   F[1631] := 3.685619;
   F[1632] := 3.6892362;
   F[1633] := 3.725405;
   F[1634] := 3.6639178;
   F[1635] := 3.6385996;
   F[1636] := 3.5879629;
   F[1637] := 3.6385996;
   F[1638] := 3.5807292;
   F[1639] := 3.59158;
   F[1640] := 3.5264757;
   F[1641] := 3.5083911;
   F[1642] := 3.5228589;
   F[1643] := 3.5300925;
   F[1644] := 3.4975405;
   F[1645] := 3.5011575;
   F[1646] := 3.4324362;
   F[1647] := 3.4252026;
   F[1648] := 3.5011575;
   F[1649] := 3.4324362;
   F[1650] := 3.410735;
   F[1651] := 3.4360533;
   F[1652] := 3.3962674;
   F[1653] := 3.374566;
   F[1654] := 3.370949;
   F[1655] := 3.3673322;
   F[1656] := 3.3528645;
   F[1657] := 3.3166957;
   F[1658] := 3.378183;
   F[1659] := 3.302228;
   F[1660] := 3.2841434;
   F[1661] := 3.294994;
   F[1662] := 3.233507;
   F[1663] := 3.2732928;
   F[1664] := 3.2045717;
   F[1665] := 3.226273;
   F[1666] := 3.1864872;
   F[1667] := 3.2045717;
   F[1668] := 3.2118056;
   F[1669] := 3.1394675;
   F[1670] := 3.157552;
   F[1671] := 3.161169;
   F[1672] := 3.1358507;
   F[1673] := 3.1286168;
   F[1674] := 3.1286168;
   F[1675] := 3.0454283;
   F[1676] := 3.0635128;
   F[1677] := 3.0996816;
   F[1678] := 3.0454283;
   F[1679] := 3.049045;
   F[1680] := 3.049045;
   F[1681] := 3.023727;
   F[1682] := 3.0092592;
   F[1683] := 2.9513888;
   F[1684] := 2.9513888;
   F[1685] := 2.983941;
   F[1686] := 2.980324;
   F[1687] := 2.9296875;
   F[1688] := 2.911603;
   F[1689] := 2.8573496;
   F[1690] := 2.8645833;
   F[1691] := 2.9188368;
   F[1692] := 2.911603;
   F[1693] := 2.8175638;
   F[1694] := 2.8537326;
   F[1695] := 2.842882;
   F[1696] := 2.8320312;
   F[1697] := 2.7958622;
   F[1698] := 2.7777777;
   F[1699] := 2.8139467;
   F[1700] := 2.734375;
   F[1701] := 2.7199075;
   F[1702] := 2.7596934;
   F[1703] := 2.7162905;
   F[1704] := 2.698206;
   F[1705] := 2.7416089;
   F[1706] := 2.6945891;
   F[1707] := 2.6801214;
   F[1708] := 2.6728878;
   F[1709] := 2.6367188;
   F[1710] := 2.629485;
   F[1711] := 2.6801214;
   F[1712] := 2.6367188;
   F[1713] := 2.6150174;
   F[1714] := 2.5752316;
   F[1715] := 2.564381;
   F[1716] := 2.55353;
   F[1717] := 2.5788484;
   F[1718] := 2.5426793;
   F[1719] := 2.4920428;
   F[1720] := 2.5282118;
   F[1721] := 2.5065105;
   F[1722] := 2.5028934;
   F[1723] := 2.4775753;
   F[1724] := 2.44864;
   F[1725] := 2.4088542;
   F[1726] := 2.4233217;
   F[1727] := 2.5065105;
   F[1728] := 2.3980036;
   F[1729] := 2.445023;
   F[1730] := 2.3582175;
   F[1731] := 2.4233217;
   F[1732] := 2.3618345;
   F[1733] := 2.376302;
   F[1734] := 2.3654513;
   F[1735] := 2.2858796;
   F[1736] := 2.3184316;
   F[1737] := 2.23886;
   F[1738] := 2.3365161;
   F[1739] := 2.275029;
   F[1740] := 2.2605612;
   F[1741] := 2.1918402;
   F[1742] := 2.2280092;
   F[1743] := 1.634838;
   F[1744] := 0.9765625;
   F[1745] := 0.30020255;
   F[1746] := 3.4432871;
   F[1747] := 5.0455728;
   F[1748] := 5.0998263;
   F[1749] := 5.10706;
   F[1750] := 5.0853586;
   F[1751] := 5.1613135;
   F[1752] := 5.117911;
   F[1753] := 5.128762;
   F[1754] := 5.0925927;
   F[1755] := 5.143229;
   F[1756] := 5.0600405;
   F[1757] := 5.0708914;
   F[1758] := 5.1649303;
   F[1759] := 5.128762;
   F[1760] := 5.114294;
   F[1761] := 5.103443;
   F[1762] := 5.1576967;
   F[1763] := 5.183015;
   F[1764] := 5.117911;
   F[1765] := 5.1576967;
   F[1766] := 5.179398;
   F[1767] := 5.1649303;
   F[1768] := 5.0708914;
   F[1769] := 5.1251445;
   F[1770] := 5.215567;
   F[1771] := 5.179398;
   F[1772] := 5.2119503;
   F[1773] := 5.1721644;
   F[1774] := 5.204716;
   F[1775] := 5.150463;
   F[1776] := 5.204716;
   F[1777] := 5.179398;
   F[1778] := 5.190249;
   F[1779] := 5.1974826;
   F[1780] := 5.2445025;
   F[1781] := 5.2408853;
   F[1782] := 5.1757812;
   F[1783] := 5.251736;
   F[1784] := 5.280671;
   F[1785] := 5.2445025;
   F[1786] := 5.255353;
   F[1787] := 5.2842884;
   F[1788] := 5.2408853;
   F[1789] := 5.280671;
   F[1790] := 5.2445025;
   F[1791] := 5.2336516;
   F[1792] := 5.2987556;
   F[1793] := 5.230035;
   F[1794] := 5.2698207;
   F[1795] := 5.31684;
   F[1796] := 5.3783274;
   F[1797] := 5.3385415;
   F[1798] := 5.2987556;
   F[1799] := 5.287905;
   F[1800] := 5.3132234;
   F[1801] := 5.2770543;
   F[1802] := 5.3747106;
   F[1803] := 5.3132234;
   F[1804] := 5.4000287;
   F[1805] := 5.353009;
   F[1806] := 5.3096066;
   F[1807] := 5.6315103;
   F[1808] := 6.3368053;
   F[1809] := 6.969763;
   F[1810] := 7.60272;
   F[1811] := 8.282697;
   F[1812] := 8.427373;
   F[1813] := 8.405671;
   F[1814] := 8.445457;
   F[1815] := 8.456307;
   F[1816] := 8.423756;
   F[1817] := 8.510561;
   F[1818] := 8.539496;
   F[1819] := 8.564815;
   F[1820] := 8.496094;
   F[1821] := 8.59375;
   F[1822] := 8.600984;
   F[1823] := 8.619068;
   F[1824] := 8.557581;
   F[1825] := 8.691406;
   F[1826] := 8.669704;
   F[1827] := 8.691406;
   F[1828] := 8.738426;
   F[1829] := 8.637153;
   F[1830] := 8.763744;
   F[1831] := 8.781829;
   F[1832] := 8.796296;
   F[1833] := 8.785445;
   F[1834] := 8.80353;
   F[1835] := 8.843316;
   F[1836] := 8.854167;
   F[1837] := 8.875868;
   F[1838] := 8.843316;
   F[1839] := 8.908421;
   F[1840] := 8.937355;
   F[1841] := 8.9192705;
   F[1842] := 9.006077;
   F[1843] := 8.959057;
   F[1844] := 8.998842;
   F[1845] := 8.973524;
   F[1846] := 9.016927;
   F[1847] := 9.031395;
   F[1848] := 9.031395;
   F[1849] := 8.998842;
   F[1850] := 9.085649;
   F[1851] := 9.063947;
   F[1852] := 9.154369;
   F[1853] := 9.186921;
   F[1854] := 9.161603;
   F[1855] := 9.273726;
   F[1856] := 9.201389;
   F[1857] := 9.226707;
   F[1858] := 9.233941;
   F[1859] := 9.248408;
   F[1860] := 9.248408;
   F[1861] := 9.338831;
   F[1862] := 9.338831;
   F[1863] := 9.349682;
   F[1864] := 9.302662;
   F[1865] := 9.364149;
   F[1866] := 9.447338;
   F[1867] := 9.367766;
   F[1868] := 9.454572;
   F[1869] := 9.385851;
   F[1870] := 9.42202;
   F[1871] := 9.476274;
   F[1872] := 9.490741;
   F[1873] := 9.505208;
   F[1874] := 9.505208;
   F[1875] := 9.602864;
   F[1876] := 9.555845;
   F[1877] := 9.544994;
   F[1878] := 9.588397;
   F[1879] := 9.628182;
   F[1880] := 9.664351;
   F[1881] := 9.628182;
   F[1882] := 9.660735;
   F[1883] := 9.682436;
   F[1884] := 9.729456;
   F[1885] := 9.707755;
   F[1886] := 9.73669;
   F[1887] := 9.740307;
   F[1888] := 9.823495;
   F[1889] := 9.805411;
   F[1890] := 9.798177;
   F[1891] := 9.823495;
   F[1892] := 9.866899;
   F[1893] := 9.881366;
   F[1894] := 9.85243;
   F[1895] := 9.975405;
   F[1896] := 10.007957;
   F[1897] := 9.95732;
   F[1898] := 10.029658;
   F[1899] := 10.185185;
   F[1900] := 10.206886;
   F[1901] := 10.315393;
   F[1902] := 10.467303;
   F[1903] := 10.554109;
   F[1904] := 10.691551;
   F[1905] := 10.756655;
   F[1906] := 10.789207;
   F[1907] := 10.966435;
   F[1908] := 11.067708;
   F[1909] := 11.161748;
   F[1910] := 11.205151;
   F[1911] := 11.338976;
   F[1912] := 11.472801;
   F[1913] := 11.555989;
   F[1914] := 11.603009;
   F[1915] := 11.715133;
   F[1916] := 11.794704;
   F[1917] := 11.924913;
   F[1918] := 12.040654;
   F[1919] := 12.131077;
   F[1920] := 12.203414;
   F[1921] := 12.355324;
   F[1922] := 12.384259;
   F[1923] := 12.507234;
   F[1924] := 12.60489;
   F[1925] := 12.648293;
   F[1926] := 12.800202;
   F[1927] := 12.9557295;
   F[1928] := 13.042535;
   F[1929] := 13.078704;
   F[1930] := 13.165509;
   F[1931] := 13.32827;
   F[1932] := 13.404224;
   F[1933] := 13.527199;
   F[1934] := 13.58507;
   F[1935] := 13.726129;
   F[1936] := 13.820168;
   F[1937] := 13.968461;
   F[1938] := 13.990162;
   F[1939] := 14.134838;
   F[1940] := 14.21441;
   F[1941] := 14.279514;
   F[1942] := 14.362702;
   F[1943] := 14.532697;
   F[1944] := 14.619502;
   F[1945] := 14.7316265;
   F[1946] := 14.840133;
   F[1947] := 14.923322;
   F[1948] := 14.623119;
   F[1949] := 13.798467;
   F[1950] := 12.9557295;
   F[1951] := 12.160011;
   F[1952] := 11.382379;
   F[1953] := 11.020689;
   F[1954] := 11.053241;
   F[1955] := 11.121962;
   F[1956] := 11.107494;
   F[1957] := 11.143663;
   F[1958] := 11.121962;
   F[1959] := 11.150897;
   F[1960] := 11.14728;
   F[1961] := 11.219618;
   F[1962] := 11.190682;
   F[1963] := 11.183449;
   F[1964] := 11.223235;
   F[1965] := 11.302807;
   F[1966] := 11.295573;
   F[1967] := 11.255787;
   F[1968] := 11.364294;
   F[1969] := 11.317274;
   F[1970] := 11.375145;
   F[1971] := 11.3932295;
   F[1972] := 11.418548;
   F[1973] := 11.4402485;
   F[1974] := 11.469184;
   F[1975] := 11.436632;
   F[1976] := 11.494502;
   F[1977] := 11.494502;
   F[1978] := 11.588542;
   F[1979] := 11.555989;
   F[1980] := 11.559607;
   F[1981] := 11.603009;
   F[1982] := 11.617476;
   F[1983] := 11.617476;
   F[1984] := 11.704283;
   F[1985] := 11.693432;
   F[1986] := 11.678964;
   F[1987] := 11.715133;
   F[1988] := 11.744068;
   F[1989] := 11.773004;
   F[1990] := 11.758536;
   F[1991] := 11.816406;
   F[1992] := 11.809173;
   F[1993] := 11.848958;
   F[1994] := 11.910445;
   F[1995] := 11.950232;
   F[1996] := 11.874276;
   F[1997] := 11.932147;
   F[1998] := 11.924913;
   F[1999] := 11.968316;
   F[2000] := 11.979167;
   F[2001] := 12.004485;
   F[2002] := 12.037037;
   F[2003] := 12.000868;
   F[2004] := 12.123842;
   F[2005] := 12.105758;
   F[2006] := 12.181713;
   F[2007] := 12.141927;
   F[2008] := 12.203414;
   F[2009] := 12.13831;
   F[2010] := 12.203414;
   F[2011] := 12.239583;
   F[2012] := 12.250434;
   F[2013] := 12.2432;
   F[2014] := 12.29022;
   F[2015] := 12.326389;
   F[2016] := 12.366175;
   F[2017] := 12.362557;
   F[2018] := 12.358941;
   F[2019] := 12.3878765;
   F[2020] := 12.3878765;
   F[2021] := 12.424046;
   F[2022] := 12.405961;
   F[2023] := 12.485533;
   F[2024] := 12.528935;
   F[2025] := 12.528935;
   F[2026] := 12.528935;
   F[2027] := 12.54702;
   F[2028] := 12.554254;
   F[2029] := 12.615741;
   F[2030] := 12.619358;
   F[2031] := 12.626592;
   F[2032] := 12.662761;
   F[2033] := 12.6953125;
   F[2034] := 12.764033;
   F[2035] := 12.811053;
   F[2036] := 12.724248;
   F[2037] := 12.760417;
   F[2038] := 12.80382;
   F[2039] := 12.843605;
   F[2040] := 12.836371;
   F[2041] := 12.850839;
   F[2042] := 12.90871;
   F[2043] := 12.941261;
   F[2044] := 13.292101;
   F[2045] := 15.704572;
   F[2046] := 18.17853;
   F[2047] := 20.706741;
   F[2048] := 23.1807;
   F[2049] := 25.672743;
   F[2050] := 28.121384;
   F[2051] := 30.671297;
   F[2052] := 33.15249;
   F[2053] := 35.633682;
   F[2054] := 38.151043;
   F[2055] := 40.588833;
   F[2056] := 40.559895;
   F[2057] := 37.492767;
   F[2058] := 34.964554;
   F[2059] := 32.508682;
   F[2060] := 30.016638;
   F[2061] := 27.50651;
   F[2062] := 25.043404;
   F[2063] := 22.518808;
   F[2064] := 20.070168;
   F[2065] := 17.520254;
   F[2066] := 15.089699;
   F[2067] := 12.579572;
   F[2068] := 11.237702;
   F[2069] := 11.161748;
   F[2070] := 11.2160015;
   F[2071] := 11.114728;
   F[2072] := 11.100261;
   F[2073] := 11.121962;
   F[2074] := 11.096643;
   F[2075] := 11.085793;
   F[2076] := 11.031539;
   F[2077] := 11.024305;
   F[2078] := 11.056858;
   F[2079] := 10.951967;
   F[2080] := 11.020689;
   F[2081] := 10.944734;
   F[2082] := 10.912182;
   F[2083] := 10.901331;
   F[2084] := 10.87963;
   F[2085] := 10.8253765;
   F[2086] := 10.803675;
   F[2087] := 10.789207;
   F[2088] := 10.73857;
   F[2089] := 10.745805;
   F[2090] := 10.781974;
   F[2091] := 10.706018;
   F[2092] := 10.724103;
   F[2093] := 10.593895;
   F[2094] := 10.673467;
   F[2095] := 10.6807;
   F[2096] := 10.572193;
   F[2097] := 10.554109;
   F[2098] := 10.579427;
   F[2099] := 10.503472;
   F[2100] := 10.521557;
   F[2101] := 10.52879;
   F[2102] := 10.463686;
   F[2103] := 10.445601;
   F[2104] := 10.46007;
   F[2105] := 10.532408;
   F[2106] := 10.420283;
   F[2107] := 10.35518;
   F[2108] := 10.322627;
   F[2109] := 10.326244;
   F[2110] := 10.3515625;
   F[2111] := 10.286458;
   F[2112] := 10.250289;
   F[2113] := 10.243055;
   F[2114] := 10.228588;
   F[2115] := 10.2213545;
   F[2116] := 10.181568;
   F[2117] := 10.206886;
   F[2118] := 10.192419;
   F[2119] := 10.083912;
   F[2120] := 10.112847;
   F[2121] := 10.083912;
   F[2122] := 10.054976;
   F[2123] := 10.047743;
   F[2124] := 10.007957;
   F[2125] := 10.007957;
   F[2126] := 9.964555;
   F[2127] := 9.982639;
   F[2128] := 9.986256;
   F[2129] := 9.924768;
   F[2130] := 9.89945;
   F[2131] := 9.892217;
   F[2132] := 9.848814;
   F[2133] := 9.837963;
   F[2134] := 9.884983;
   F[2135] := 9.801794;
   F[2136] := 9.780092;
   F[2137] := 9.780092;
   F[2138] := 9.754774;
   F[2139] := 9.725839;
   F[2140] := 9.725839;
   F[2141] := 9.711371;
   F[2142] := 9.693287;
   F[2143] := 9.6535015;
   F[2144] := 9.617332;
   F[2145] := 9.628182;
   F[2146] := 9.599248;
   F[2147] := 9.566695;
   F[2148] := 9.610099;
   F[2149] := 9.57393;
   F[2150] := 9.508825;
   F[2151] := 9.4871235;
   F[2152] := 9.443721;
   F[2153] := 9.414786;
   F[2154] := 9.43287;
   F[2155] := 9.382234;
   F[2156] := 9.382234;
   F[2157] := 9.360533;
   F[2158] := 9.324364;
   F[2159] := 9.338831;
   F[2160] := 9.306279;
   F[2161] := 9.378617;
   F[2162] := 9.244792;
   F[2163] := 9.215857;
   F[2164] := 9.2628765;
   F[2165] := 9.291811;
   F[2166] := 9.186921;
   F[2167] := 9.183305;
   F[2168] := 9.190538;
   F[2169] := 9.194155;
   F[2170] := 9.147136;
   F[2171] := 9.067564;
   F[2172] := 9.035011;
   F[2173] := 9.009693;
   F[2174] := 9.103733;
   F[2175] := 8.991609;
   F[2176] := 9.009693;
   F[2177] := 9.009693;
   F[2178] := 8.991609;
   F[2179] := 9.027778;
   F[2180] := 8.933739;
   F[2181] := 8.8722515;
   F[2182] := 8.933739;
   F[2183] := 8.865017;
   F[2184] := 8.875868;
   F[2185] := 8.843316;
   F[2186] := 8.7890625;
   F[2187] := 8.843316;
   F[2188] := 8.74566;
   F[2189] := 8.713108;
   F[2190] := 8.767361;
   F[2191] := 8.7058735;
   F[2192] := 8.687789;
   F[2193] := 8.673322;
   F[2194] := 8.7058735;
   F[2195] := 8.600984;
   F[2196] := 8.597367;
   F[2197] := 8.604601;
   F[2198] := 8.600984;
   F[2199] := 8.575665;
   F[2200] := 8.532263;
   F[2201] := 8.532263;
   F[2202] := 8.521412;
   F[2203] := 8.553964;
   F[2204] := 8.5286455;
   F[2205] := 8.478009;
   F[2206] := 8.4816265;
   F[2207] := 8.470776;
   F[2208] := 8.409288;
   F[2209] := 8.351418;
   F[2210] := 8.308015;
   F[2211] := 8.362268;
   F[2212] := 8.3152485;
   F[2213] := 8.3152485;
   F[2214] := 8.297164;
   F[2215] := 8.293548;
   F[2216] := 8.213976;
   F[2217] := 8.206742;
   F[2218] := 8.199508;
   F[2219] := 8.224827;
   F[2220] := 8.192274;
   F[2221] := 8.17419;
   F[2222] := 8.18504;
   F[2223] := 8.134404;
   F[2224] := 8.101851;
   F[2225] := 8.065682;
   F[2226] := 8.080151;
   F[2227] := 8.065682;
   F[2228] := 8.065682;
   F[2229] := 8.025897;
   F[2230] := 7.9716434;
   F[2231] := 8.036748;
   F[2232] := 7.9318576;
   F[2233] := 7.939091;
   F[2234] := 7.949942;
   F[2235] := 7.913773;
   F[2236] := 7.9029226;
   F[2237] := 7.8703704;
   F[2238] := 7.884838;
   F[2239] := 7.8956885;
   F[2240] := 7.837818;
   F[2241] := 7.8052664;
   F[2242] := 7.747396;
   F[2243] := 7.7582464;
   F[2244] := 7.7256947;
   F[2245] := 7.7546296;
   F[2246] := 7.703993;
   F[2247] := 7.6931424;
   F[2248] := 7.7293115;
   F[2249] := 7.6678243;
   F[2250] := 7.6171875;
   F[2251] := 7.5882525;
   F[2252] := 7.6497397;
   F[2253] := 7.5810184;
   F[2254] := 7.573785;
   F[2255] := 7.5810184;
   F[2256] := 7.530382;
   F[2257] := 7.5520835;
   F[2258] := 7.5050635;
   F[2259] := 7.486979;
   F[2260] := 7.472512;
   F[2261] := 7.5014467;
   F[2262] := 7.396557;
   F[2263] := 7.382089;
   F[2264] := 7.458044;
   F[2265] := 7.360388;
   F[2266] := 7.3423033;
   F[2267] := 7.349537;
   F[2268] := 7.309751;
   F[2269] := 7.3025174;
   F[2270] := 7.248264;
   F[2271] := 7.306134;
   F[2272] := 7.269965;
   F[2273] := 7.2265625;
   F[2274] := 7.1903934;
   F[2275] := 7.157841;
   F[2276] := 7.2012444;
   F[2277] := 7.139757;
   F[2278] := 7.168692;
   F[2279] := 7.1108217;
   F[2280] := 7.081887;
   F[2281] := 7.0746527;
   F[2282] := 7.0999713;
   F[2283] := 7.0457177;
   F[2284] := 7.1759257;
   F[2285] := 7.027633;
   F[2286] := 7.03125;
   F[2287] := 6.9878473;
   F[2288] := 6.9733796;
   F[2289] := 7.0131655;
   F[2290] := 6.929977;
   F[2291] := 6.8757234;
   F[2292] := 6.8974247;
   F[2293] := 6.857639;
   F[2294] := 6.8467884;
   F[2295] := 6.8865743;
   F[2296] := 6.8106194;
   F[2297] := 6.7599826;
   F[2298] := 6.792535;
   F[2299] := 6.814236;
   F[2300] := 6.792535;
   F[2301] := 6.2970195;
   F[2302] := 5.6351275;
   F[2303] := 4.875579;
   F[2304] := 4.257089;
   F[2305] := 3.6639178;
   F[2306] := 3.7073207;
   F[2307] := 3.69647;
   F[2308] := 3.6385996;
   F[2309] := 3.692853;
   F[2310] := 3.685619;
   F[2311] := 3.660301;
   F[2312] := 3.6639178;
   F[2313] := 3.6385996;
   F[2314] := 3.656684;
   F[2315] := 3.7181714;
   F[2316] := 3.685619;
   F[2317] := 3.6422164;
   F[2318] := 3.6277487;
   F[2319] := 3.620515;
   F[2320] := 3.6458333;
   F[2321] := 3.6385996;
   F[2322] := 3.5951967;
   F[2323] := 3.584346;
   F[2324] := 3.6313658;
   F[2325] := 3.5988138;
   F[2326] := 3.5879629;
   F[2327] := 3.5807292;
   F[2328] := 3.5879629;
   F[2329] := 3.5554109;
   F[2330] := 3.5879629;
   F[2331] := 3.59158;
   F[2332] := 3.551794;
   F[2333] := 3.5300925;
   F[2334] := 3.6060474;
   F[2335] := 3.5554109;
   F[2336] := 3.5300925;
   F[2337] := 3.5409434;
   F[2338] := 3.5264757;
   F[2339] := 3.5047743;
   F[2340] := 3.5192418;
   F[2341] := 3.5083911;
   F[2342] := 3.5373263;
   F[2343] := 3.5626447;
   F[2344] := 3.5011575;
   F[2345] := 3.5409434;
   F[2346] := 3.4866898;
   F[2347] := 3.5662615;
   F[2348] := 3.5120082;
   F[2349] := 3.5047743;
   F[2350] := 3.5192418;
   F[2351] := 3.4903066;
   F[2352] := 3.5228589;
   F[2353] := 3.4866898;
   F[2354] := 3.4505208;
   F[2355] := 3.4722223;
   F[2356] := 3.4649885;
   F[2357] := 3.446904;
   F[2358] := 3.4577546;
   F[2359] := 3.3528645;
   F[2360] := 3.4939237;
   F[2361] := 3.4866898;
   F[2362] := 3.4179688;
   F[2363] := 3.4215856;
   F[2364] := 3.4252026;
   F[2365] := 3.378183;
   F[2366] := 1.8916377;
   F[2367] := 4.615162;
   F[2368] := 4.626013;
   F[2369] := 4.5645256;
   F[2370] := 4.6187787;
   F[2371] := 4.6187787;
   F[2372] := 4.560909;
   F[2373] := 4.662182;
   F[2374] := 4.6296296;
   F[2375] := 4.6187787;
   F[2376] := 4.615162;
   F[2377] := 4.5645256;
   F[2378] := 4.622396;
   F[2379] := 4.6079283;
   F[2380] := 4.658565;
   F[2381] := 4.683883;
   F[2382] := 4.622396;
   F[2383] := 4.6043115;
   F[2384] := 4.691117;
   F[2385] := 4.6875;
   F[2386] := 4.676649;
   F[2387] := 4.647714;
   F[2388] := 4.6440973;
   F[2389] := 4.651331;
   F[2390] := 4.691117;
   F[2391] := 4.5898438;
   F[2392] := 4.6043115;
   F[2393] := 4.6730323;
   F[2394] := 4.723669;
   F[2395] := 4.6332464;
   F[2396] := 4.6730323;
   F[2397] := 4.7019677;
   F[2398] := 4.727286;
   F[2399] := 4.698351;
   F[2400] := 4.7019677;
   F[2401] := 4.6875;
   F[2402] := 4.6802664;
   F[2403] := 4.6730323;
   F[2404] := 4.6802664;
   F[2405] := 4.716435;
   F[2406] := 4.6947336;
   F[2407] := 4.6549478;
   F[2408] := 4.727286;
   F[2409] := 4.7345195;
   F[2410] := 4.738137;
   F[2411] := 4.727286;
   F[2412] := 4.788773;
   F[2413] := 4.7815394;
   F[2414] := 4.788773;
   F[2415] := 4.7670717;
   F[2416] := 4.7706885;
   F[2417] := 4.799624;
   F[2418] := 4.738137;
   F[2419] := 4.738137;
   F[2420] := 4.8177085;
   F[2421] := 4.763455;
   F[2422] := 4.8574944;
   F[2423] := 4.7815394;
   F[2424] := 4.7670717;
   F[2425] := 4.796007;
   F[2426] := 4.803241;
   F[2427] := 4.9479165;
   F[2428] := 5.5917244;
   F[2429] := 6.2934027;
   F[2430] := 6.919126;
   F[2431] := 7.526765;
   F[2432] := 7.8956885;
   F[2433] := 7.8920717;
   F[2434] := 7.8920717;
   F[2435] := 7.939091;
   F[2436] := 7.9029226;
   F[2437] := 7.960793;
   F[2438] := 7.960793;
   F[2439] := 7.960793;
   F[2440] := 7.9788775;
   F[2441] := 7.96441;
   F[2442] := 7.9463253;
   F[2443] := 8.036748;
   F[2444] := 8.018663;
   F[2445] := 8.087384;
   F[2446] := 8.065682;
   F[2447] := 8.105469;
   F[2448] := 8.141638;
   F[2449] := 8.188658;
   F[2450] := 8.145255;
   F[2451] := 8.181423;
   F[2452] := 8.192274;
   F[2453] := 8.17419;
   F[2454] := 8.275463;
   F[2455] := 8.206742;
   F[2456] := 8.199508;
   F[2457] := 8.308015;
   F[2458] := 8.257379;
   F[2459] := 8.311632;
   F[2460] := 8.326099;
   F[2461] := 8.33695;
   F[2462] := 8.322483;
   F[2463] := 8.33695;
   F[2464] := 8.3152485;
   F[2465] := 8.412905;
   F[2466] := 8.380353;
   F[2467] := 8.344184;
   F[2468] := 8.463542;
   F[2469] := 8.412905;
   F[2470] := 8.467158;
   F[2471] := 8.459925;
   F[2472] := 8.525029;
   F[2473] := 8.496094;
   F[2474] := 8.499711;
   F[2475] := 8.568432;
   F[2476] := 8.499711;
   F[2477] := 8.575665;
   F[2478] := 8.564815;
   F[2479] := 8.619068;
   F[2480] := 8.626302;
   F[2481] := 8.684173;
   F[2482] := 8.629919;
   F[2483] := 8.684173;
   F[2484] := 8.69864;
   F[2485] := 8.662471;
   F[2486] := 8.713108;
   F[2487] := 8.716724;
   F[2488] := 8.785445;
   F[2489] := 8.774595;
   F[2490] := 8.785445;
   F[2491] := 8.7890625;
   F[2492] := 8.79268;
   F[2493] := 8.846932;
   F[2494] := 8.825232;
   F[2495] := 8.904803;
   F[2496] := 8.890336;
   F[2497] := 8.930121;
   F[2498] := 8.987992;
   F[2499] := 8.973524;
   F[2500] := 8.944589;
   F[2501] := 8.933739;
   F[2502] := 9.07118;
   F[2503] := 9.01331;
   F[2504] := 9.038629;
   F[2505] := 9.020544;
   F[2506] := 9.056713;
   F[2507] := 9.07118;
   F[2508] := 9.038629;
   F[2509] := 9.125434;
   F[2510] := 9.1182;
   F[2511] := 9.103733;
   F[2512] := 9.190538;
   F[2513] := 9.139901;
   F[2514] := 9.215857;
   F[2515] := 9.244792;
   F[2516] := 9.226707;
   F[2517] := 9.284577;
   F[2518] := 9.302662;
   F[2519] := 9.400318;
   F[2520] := 9.519676;
   F[2521] := 9.602864;
   F[2522] := 9.696904;
   F[2523] := 9.801794;
   F[2524] := 9.870515;
   F[2525] := 9.94647;
   F[2526] := 10.058594;
   F[2527] := 10.174335;
   F[2528] := 10.275608;
   F[2529] := 10.380498;
   F[2530] := 10.456452;
   F[2531] := 10.568577;
   F[2532] := 10.698785;
   F[2533] := 10.745805;
   F[2534] := 10.836226;
   F[2535] := 10.944734;
   F[2536] := 11.078559;
   F[2537] := 11.085793;
   F[2538] := 11.248553;
   F[2539] := 11.367911;
   F[2540] := 11.458333;
   F[2541] := 11.530671;
   F[2542] := 11.621094;
   F[2543] := 11.700665;
   F[2544] := 11.841724;
   F[2545] := 11.92853;
   F[2546] := 12.029803;
   F[2547] := 12.152778;
   F[2548] := 12.207031;
   F[2549] := 12.344474;
   F[2550] := 12.377026;
   F[2551] := 12.518085;
   F[2552] := 12.637443;
   F[2553] := 12.713397;
   F[2554] := 12.811053;
   F[2555] := 12.883391;
   F[2556] := 13.064236;
   F[2557] := 13.089555;
   F[2558] := 13.22338;
   F[2559] := 13.292101;
   F[2560] := 13.436776;
   F[2561] := 13.527199;
   F[2562] := 13.610388;
   F[2563] := 13.718895;
   F[2564] := 13.820168;
   F[2565] := 13.932292;
   F[2566] := 14.001013;
   F[2567] := 14.073351;
   F[2568] := 13.943142;
   F[2569] := 13.136574;
   F[2570] := 12.380642;
   F[2571] := 11.563224;
   F[2572] := 10.662616;
   F[2573] := 10.199653;
   F[2574] := 10.206886;
   F[2575] := 10.275608;
   F[2576] := 10.264757;
   F[2577] := 10.257524;
   F[2578] := 10.271991;
   F[2579] := 10.282842;
   F[2580] := 10.322627;
   F[2581] := 10.402199;
   F[2582] := 10.3515625;
   F[2583] := 10.36603;
   F[2584] := 10.423901;
   F[2585] := 10.470921;
   F[2586] := 10.489005;
   F[2587] := 10.478154;
   F[2588] := 10.536024;
   F[2589] := 10.525173;
   F[2590] := 10.521557;
   F[2591] := 10.539641;
   F[2592] := 10.568577;
   F[2593] := 10.622829;
   F[2594] := 10.604745;
   F[2595] := 10.640914;
   F[2596] := 10.63368;
   F[2597] := 10.615596;
   F[2598] := 10.6589985;
   F[2599] := 10.698785;
   F[2600] := 10.767506;
   F[2601] := 10.687934;
   F[2602] := 10.724103;
   F[2603] := 10.78559;
   F[2604] := 10.807292;
   F[2605] := 10.854311;
   F[2606] := 10.756655;
   F[2607] := 10.821759;
   F[2608] := 10.774739;
   F[2609] := 10.876013;
   F[2610] := 10.857928;
   F[2611] := 10.894097;
   F[2612] := 10.857928;
   F[2613] := 10.926649;
   F[2614] := 10.930266;
   F[2615] := 10.988136;
   F[2616] := 11.035156;
   F[2617] := 11.046007;
   F[2618] := 11.038774;
   F[2619] := 11.017072;
   F[2620] := 11.096643;
   F[2621] := 11.118345;
   F[2622] := 11.085793;
   F[2623] := 11.143663;
   F[2624] := 11.201533;
   F[2625] := 11.1943;
   F[2626] := 11.201533;
   F[2627] := 11.176215;
   F[2628] := 11.230469;
   F[2629] := 11.205151;
   F[2630] := 11.342592;
   F[2631] := 11.291956;
   F[2632] := 11.31004;
   F[2633] := 11.313658;
   F[2634] := 11.313658;
   F[2635] := 11.331742;
   F[2636] := 11.41493;
   F[2637] := 11.443866;
   F[2638] := 11.407697;
   F[2639] := 11.46195;
   F[2640] := 11.447483;
   F[2641] := 11.490886;
   F[2642] := 11.51982;
   F[2643] := 11.541522;
   F[2644] := 11.545139;
   F[2645] := 11.501736;
   F[2646] := 11.628327;
   F[2647] := 11.621094;
   F[2648] := 11.628327;
   F[2649] := 11.639178;
   F[2650] := 11.624711;
   F[2651] := 11.646412;
   F[2652] := 11.682581;
   F[2653] := 11.729601;
   F[2654] := 11.71875;
   F[2655] := 11.791088;
   F[2656] := 11.794704;
   F[2657] := 11.856193;
   F[2658] := 11.834491;
   F[2659] := 11.780237;
   F[2660] := 11.845342;
   F[2661] := 11.852575;
   F[2662] := 11.859809;
   F[2663] := 11.932147;
   F[2664] := 12.084057;
   F[2665] := 14.369936;
   F[2666] := 16.880064;
   F[2667] := 19.382957;
   F[2668] := 21.849682;
   F[2669] := 24.374277;
   F[2670] := 26.837385;
   F[2671] := 29.394531;
   F[2672] := 31.807003;
   F[2673] := 34.324364;
   F[2674] := 36.816406;
   F[2675] := 39.304832;
   F[2676] := 41.82581;
   F[2677] := 41.822193;
   F[2678] := 38.697193;
   F[2679] := 36.23047;
   F[2680] := 33.716724;
   F[2681] := 31.210215;
   F[2682] := 28.68562;
   F[2683] := 26.182726;
   F[2684] := 23.672598;
   F[2685] := 21.216724;
   F[2686] := 18.75;
   F[2687] := 16.26519;
   F[2688] := 13.75868;
   F[2689] := 11.2160015;
   F[2690] := 10.21412;
   F[2691] := 10.170717;
   F[2692] := 10.199653;
   F[2693] := 10.116464;
   F[2694] := 10.058594;
   F[2695] := 10.112847;
   F[2696] := 10.073061;
   F[2697] := 10.10923;
   F[2698] := 10.080296;
   F[2699] := 9.993489;
   F[2700] := 10.015191;
   F[2701] := 10.040509;
   F[2702] := 9.968171;
   F[2703] := 9.928386;
   F[2704] := 9.924768;
   F[2705] := 9.982639;
   F[2706] := 9.942853;
   F[2707] := 9.859664;
   F[2708] := 9.870515;
   F[2709] := 9.845197;
   F[2710] := 9.845197;
   F[2711] := 9.834346;
   F[2712] := 9.85243;
   F[2713] := 9.686053;
   F[2714] := 9.765625;
   F[2715] := 9.725839;
   F[2716] := 9.73669;
   F[2717] := 9.718605;
   F[2718] := 9.7005205;
   F[2719] := 9.671586;
   F[2720] := 9.628182;
   F[2721] := 9.613715;
   F[2722] := 9.599248;
   F[2723] := 9.508825;
   F[2724] := 9.519676;
   F[2725] := 9.508825;
   F[2726] := 9.47989;
   F[2727] := 9.530526;
   F[2728] := 9.505208;
   F[2729] := 9.4401045;
   F[2730] := 9.461805;
   F[2731] := 9.458189;
   F[2732] := 9.396702;
   F[2733] := 9.360533;
   F[2734] := 9.389467;
   F[2735] := 9.295428;
   F[2736] := 9.331597;
   F[2737] := 9.306279;
   F[2738] := 9.284577;
   F[2739] := 9.313513;
   F[2740] := 9.233941;
   F[2741] := 9.295428;
   F[2742] := 9.230324;
   F[2743] := 9.226707;
   F[2744] := 9.215857;
   F[2745] := 9.136285;
   F[2746] := 9.129051;
   F[2747] := 9.0964985;
   F[2748] := 9.1182;
   F[2749] := 9.0964985;
   F[2750] := 9.056713;
   F[2751] := 9.085649;
   F[2752] := 9.042245;
   F[2753] := 9.016927;
   F[2754] := 8.998842;
   F[2755] := 9.006077;
   F[2756] := 8.959057;
   F[2757] := 8.995226;
   F[2758] := 8.933739;
   F[2759] := 8.886719;
   F[2760] := 8.868634;
   F[2761] := 8.868634;
   F[2762] := 8.886719;
   F[2763] := 8.861401;
   F[2764] := 8.825232;
   F[2765] := 8.846932;
   F[2766] := 8.723958;
   F[2767] := 8.7890625;
   F[2768] := 8.74566;
   F[2769] := 8.716724;
   F[2770] := 8.676939;
   F[2771] := 8.64077;
   F[2772] := 8.695024;
   F[2773] := 8.65162;
   F[2774] := 8.637153;
   F[2775] := 8.648004;
   F[2776] := 8.64077;
   F[2777] := 8.615452;
   F[2778] := 8.586516;
   F[2779] := 8.568432;
   F[2780] := 8.539496;
   F[2781] := 8.539496;
   F[2782] := 8.470776;
   F[2783] := 8.532263;
   F[2784] := 8.423756;
   F[2785] := 8.430989;
   F[2786] := 8.44184;
   F[2787] := 8.365886;
   F[2788] := 8.485243;
   F[2789] := 8.344184;
   F[2790] := 8.373119;
   F[2791] := 8.304399;
   F[2792] := 8.355035;
   F[2793] := 8.3152485;
   F[2794] := 8.300781;
   F[2795] := 8.246528;
   F[2796] := 8.297164;
   F[2797] := 8.257379;
   F[2798] := 8.235677;
   F[2799] := 8.206742;
   F[2800] := 8.199508;
   F[2801] := 8.177807;
   F[2802] := 8.159722;
   F[2803] := 8.152489;
   F[2804] := 8.065682;
   F[2805] := 8.148871;
   F[2806] := 8.083767;
   F[2807] := 8.065682;
   F[2808] := 8.051215;
   F[2809] := 8.047599;
   F[2810] := 8.029514;
   F[2811] := 8.01143;
   F[2812] := 7.9824944;
   F[2813] := 7.9571757;
   F[2814] := 7.9427085;
   F[2815] := 7.921007;
   F[2816] := 7.924624;
   F[2817] := 7.888455;
   F[2818] := 7.8956885;
   F[2819] := 7.8450522;
   F[2820] := 7.816117;
   F[2821] := 7.8305845;
   F[2822] := 7.873987;
   F[2823] := 7.7944155;
   F[2824] := 7.7980323;
   F[2825] := 7.675058;
   F[2826] := 7.751013;
   F[2827] := 7.736545;
   F[2828] := 7.675058;
   F[2829] := 7.6569734;
   F[2830] := 7.7329283;
   F[2831] := 7.664207;
   F[2832] := 7.6822915;
   F[2833] := 7.624421;
   F[2834] := 7.624421;
   F[2835] := 7.599103;
   F[2836] := 7.5810184;
   F[2837] := 7.5774016;
   F[2838] := 7.533999;
   F[2839] := 7.494213;
   F[2840] := 7.548466;
   F[2841] := 7.4652777;
   F[2842] := 7.530382;
   F[2843] := 7.4905963;
   F[2844] := 7.3893228;
   F[2845] := 7.411024;
   F[2846] := 7.3676214;
   F[2847] := 7.458044;
   F[2848] := 7.411024;
   F[2849] := 7.3350697;
   F[2850] := 7.3314524;
   F[2851] := 7.313368;
   F[2852] := 7.309751;
   F[2853] := 7.3025174;
   F[2854] := 7.2663484;
   F[2855] := 7.284433;
   F[2856] := 7.2374134;
   F[2857] := 7.233796;
   F[2858] := 7.244647;
   F[2859] := 7.219329;
   F[2860] := 7.132523;
   F[2861] := 7.143374;
   F[2862] := 7.143374;
   F[2863] := 7.096354;
   F[2864] := 7.0746527;
   F[2865] := 7.1289062;
   F[2866] := 7.0638022;
   F[2867] := 7.1252894;
   F[2868] := 7.0529513;
   F[2869] := 7.0638022;
   F[2870] := 7.027633;
   F[2871] := 6.9444447;
   F[2872] := 7.0638022;
   F[2873] := 6.9769964;
   F[2874] := 6.9408274;
   F[2875] := 6.966146;
   F[2876] := 6.9625287;
   F[2877] := 6.893808;
   F[2878] := 6.9625287;
   F[2879] := 6.890191;
   F[2880] := 6.890191;
   F[2881] := 6.8721066;
   F[2882] := 6.8359375;
   F[2883] := 6.8033853;
   F[2884] := 6.7997684;
   F[2885] := 6.745515;
   F[2886] := 6.749132;
   F[2887] := 6.781684;
   F[2888] := 6.702112;
   F[2889] := 6.7853007;
   F[2890] := 6.7382812;
   F[2891] := 6.7093463;
   F[2892] := 6.6731772;
   F[2893] := 6.629774;
   F[2894] := 6.6478586;
   F[2895] := 6.589988;
   F[2896] := 6.6080728;
   F[2897] := 6.6623263;
   F[2898] := 6.604456;
   F[2899] := 6.5502024;
   F[2900] := 6.5502024;
   F[2901] := 6.528501;
   F[2902] := 6.4742475;
   F[2903] := 6.503183;
   F[2904] := 6.463397;
   F[2905] := 6.4561634;
   F[2906] := 6.430845;
   F[2907] := 6.4199944;
   F[2908] := 6.4344616;
   F[2909] := 6.488715;
   F[2910] := 6.3946757;
   F[2911] := 6.391059;
   F[2912] := 6.311487;
   F[2913] := 6.351273;
   F[2914] := 6.3187213;
   F[2915] := 6.351273;
   F[2916] := 6.3078704;
   F[2917] := 6.275318;
   F[2918] := 6.2825522;
   F[2919] := 6.300637;
   F[2920] := 6.2355323;
   F[2921] := 6.25;
   F[2922] := 6.1957464;
   F[2923] := 5.5157695;
   F[2924] := 4.9189816;
   F[2925] := 4.235388;
   F[2926] := 3.6639178;
   F[2927] := 3.1394675;
   F[2928] := 3.125;
   F[2929] := 3.125;
   F[2930] := 3.092448;
   F[2931] := 3.0996816;
   F[2932] := 3.1141493;
   F[2933] := 3.1141493;
   F[2934] := 3.1213832;
   F[2935] := 3.0743635;
   F[2936] := 3.1032987;
   F[2937] := 3.092448;
   F[2938] := 3.1141493;
   F[2939] := 3.0996816;
   F[2940] := 3.1286168;
   F[2941] := 3.0381944;
   F[2942] := 3.1177661;
   F[2943] := 3.1539352;
   F[2944] := 3.0996816;
   F[2945] := 3.0635128;
   F[2946] := 3.0779803;
   F[2947] := 3.1032987;
   F[2948] := 3.0743635;
   F[2949] := 3.0309606;
   F[2950] := 3.02011;
   F[2951] := 3.0960648;
   F[2952] := 3.0635128;
   F[2953] := 3.092448;
   F[2954] := 3.0418112;
   F[2955] := 3.0526621;
   F[2956] := 3.0454283;
   F[2957] := 3.0707464;
   F[2958] := 3.0309606;
   F[2959] := 3.0345776;
   F[2960] := 3.0273438;
   F[2961] := 3.0128763;
   F[2962] := 3.0671296;
   F[2963] := 3.0020254;
   F[2964] := 3.0418112;
   F[2965] := 3.0526621;
   F[2966] := 2.9911747;
   F[2967] := 2.983941;
   F[2968] := 3.016493;
   F[2969] := 3.0598958;
   F[2970] := 3.0598958;
   F[2971] := 3.0418112;
   F[2972] := 2.9947917;
   F[2973] := 2.9911747;
   F[2974] := 3.0020254;
   F[2975] := 3.023727;
   F[2976] := 2.9911747;
   F[2977] := 2.9947917;
   F[2978] := 3.0056424;
   F[2979] := 2.9947917;
   F[2980] := 2.9767072;
   F[2981] := 2.947772;
   F[2982] := 2.9694734;
   F[2983] := 2.9694734;
   F[2984] := 2.947772;
   F[2985] := 2.9730902;
   F[2986] := 3.023727;
   F[2987] := 0.003616898;
   F[2988] := 3.8917825;
   F[2989] := 7.8667536;
   F[2990] := 10.387732;
   F[2991] := 10.405816;
   F[2992] := 10.4347515;
   F[2993] := 10.358796;
   F[2994] := 10.4347515;
   F[2995] := 10.423901;
   F[2996] := 10.423901;
   F[2997] := 10.405816;
   F[2998] := 10.391349;
   F[2999] := 10.441985;
   F[3000] := 10.423901;
   F[3001] := 10.427517;
   F[3002] := 10.445601;
   F[3003] := 10.46007;
   F[3004] := 10.463686;
   F[3005] := 10.507089;
   F[3006] := 10.4347515;
   F[3007] := 10.427517;
   F[3008] := 10.496239;
   F[3009] := 10.456452;
   F[3010] := 10.478154;
   F[3011] := 10.463686;
   F[3012] := 10.496239;
   F[3013] := 10.496239;
   F[3014] := 10.4817705;
   F[3015] := 10.416667;
   F[3016] := 10.499855;
   F[3017] := 10.51794;
   F[3018] := 10.525173;
   F[3019] := 10.532408;
   F[3020] := 10.489005;
   F[3021] := 10.507089;
   F[3022] := 10.532408;
   F[3023] := 10.496239;
   F[3024] := 10.52879;
   F[3025] := 10.590278;
   F[3026] := 10.507089;
   F[3027] := 10.550492;
   F[3028] := 10.543258;
   F[3029] := 10.561342;
   F[3030] := 10.604745;
   F[3031] := 10.590278;
   F[3032] := 10.57581;
   F[3033] := 10.601129;
   F[3034] := 10.554109;
   F[3035] := 10.543258;
   F[3036] := 10.57581;
   F[3037] := 10.604745;
   F[3038] := 10.666233;
   F[3039] := 10.640914;
   F[3040] := 10.604745;
   F[3041] := 10.6119795;
   F[3042] := 10.622829;
   F[3043] := 10.6119795;
   F[3044] := 10.63368;
   F[3045] := 10.637298;
   F[3046] := 10.669849;
   F[3047] := 10.6589985;
   F[3048] := 10.626447;
   F[3049] := 10.6807;
   F[3050] := 10.912182;
   F[3051] := 11.490886;
   F[3052] := 12.087673;
   F[3053] := 12.807436;
   F[3054] := 13.472945;
   F[3055] := 13.718895;
   F[3056] := 13.733362;
   F[3057] := 13.75868;
   F[3058] := 13.827401;
   F[3059] := 13.834636;
   F[3060] := 13.878038;
   F[3061] := 13.8671875;
   F[3062] := 13.906974;
   F[3063] := 13.86357;
   F[3064] := 13.896123;
   F[3065] := 13.928675;
   F[3066] := 13.982928;
   F[3067] := 13.964844;
   F[3068] := 14.00463;
   F[3069] := 13.939526;
   F[3070] := 14.037182;
   F[3071] := 14.033565;
   F[3072] := 14.102286;
   F[3073] := 14.1276045;
   F[3074] := 14.080585;
   F[3075] := 14.1276045;
   F[3076] := 14.102286;
   F[3077] := 14.171007;
   F[3078] := 14.156539;
   F[3079] := 14.1746235;
   F[3080] := 14.210793;
   F[3081] := 14.221643;
   F[3082] := 14.265046;
   F[3083] := 14.239728;
   F[3084] := 14.268663;
   F[3085] := 14.279514;
   F[3086] := 14.333767;
   F[3087] := 14.297599;
   F[3088] := 14.312066;
   F[3089] := 14.355469;
   F[3090] := 14.362702;
   F[3091] := 14.406105;
   F[3092] := 14.402489;
   F[3093] := 14.409722;
   F[3094] := 14.514612;
   F[3095] := 14.48206;
   F[3096] := 14.500145;
   F[3097] := 14.510995;
   F[3098] := 14.456742;
   F[3099] := 14.525463;
   F[3100] := 14.561632;
   F[3101] := 14.63397;
   F[3102] := 14.58695;
   F[3103] := 14.615886;
   F[3104] := 14.63397;
   F[3105] := 14.688224;
   F[3106] := 14.655671;
   F[3107] := 14.670139;
   F[3108] := 14.713542;
   F[3109] := 14.709925;
   F[3110] := 14.775029;
   F[3111] := 14.782263;
   F[3112] := 14.800347;
   F[3113] := 14.811198;
   F[3114] := 14.847367;
   F[3115] := 14.9088545;
   F[3116] := 14.854601;
   F[3117] := 14.869068;
   F[3118] := 14.90162;
   F[3119] := 14.934173;
   F[3120] := 14.923322;
   F[3121] := 14.959491;
   F[3122] := 14.945024;
   F[3123] := 15.002893;
   F[3124] := 15.028212;
   F[3125] := 15.05353;
   F[3126] := 15.0390625;
   F[3127] := 15.071614;
   F[3128] := 15.060764;
   F[3129] := 15.075232;
   F[3130] := 15.143952;
   F[3131] := 15.140336;
   F[3132] := 15.165654;
   F[3133] := 15.172888;
   F[3134] := 15.194589;
   F[3135] := 15.212673;
   F[3136] := 15.237992;
   F[3137] := 15.230758;
   F[3138] := 15.274161;
   F[3139] := 15.292245;
   F[3140] := 15.259693;
   F[3141] := 15.436921;
   F[3142] := 15.47309;
   F[3143] := 15.56713;
   F[3144] := 15.704572;
   F[3145] := 15.809462;
   F[3146] := 15.925202;
   F[3147] := 15.99754;
   F[3148] := 16.040943;
   F[3149] := 16.229021;
   F[3150] := 16.29051;
   F[3151] := 16.413485;
   F[3152] := 16.45327;
   F[3153] := 16.594328;
   F[3154] := 16.735388;
   F[3155] := 16.771557;
   F[3156] := 16.945168;
   F[3157] := 16.974104;
   F[3158] := 17.086227;
   F[3159] := 17.126013;
   F[3160] := 17.256222;
   F[3161] := 17.386429;
   F[3162] := 17.520254;
   F[3163] := 17.563658;
   F[3164] := 17.690248;
   F[3165] := 17.82769;
   F[3166] := 17.914497;
   F[3167] := 17.939816;
   F[3168] := 18.051939;
   F[3169] := 18.171297;
   F[3170] := 18.254484;
   F[3171] := 18.381077;
   F[3172] := 18.525753;
   F[3173] := 18.612558;
   F[3174] := 18.663195;
   F[3175] := 18.757235;
   F[3176] := 18.898293;
   F[3177] := 18.981482;
   F[3178] := 19.089989;
   F[3179] := 19.245516;
   F[3180] := 19.288918;
   F[3181] := 19.433594;
   F[3182] := 19.560184;
   F[3183] := 19.599972;
   F[3184] := 19.62529;
   F[3185] := 19.806135;
   F[3186] := 19.896557;
   F[3187] := 19.979746;
   F[3188] := 20.120804;
   F[3189] := 20.225695;
   F[3190] := 20.330584;
   F[3191] := 20.272715;
   F[3192] := 19.480614;
   F[3193] := 18.565538;
   F[3194] := 17.856627;
   F[3195] := 17.006655;
   F[3196] := 16.485823;
   F[3197] := 16.44242;
   F[3198] := 16.550926;
   F[3199] := 16.456886;
   F[3200] := 16.540075;
   F[3201] := 16.56901;
   F[3202] := 16.554543;
   F[3203] := 16.608797;
   F[3204] := 16.597946;
   F[3205] := 16.659433;
   F[3206] := 16.71007;
   F[3207] := 16.724537;
   F[3208] := 16.735388;
   F[3209] := 16.677517;
   F[3210] := 16.728153;
   F[3211] := 16.735388;
   F[3212] := 16.861979;
   F[3213] := 16.796875;
   F[3214] := 16.83666;
   F[3215] := 16.847511;
   F[3216] := 16.854746;
   F[3217] := 16.912615;
   F[3218] := 16.876448;
   F[3219] := 16.959635;
   F[3220] := 17.006655;
   F[3221] := 16.934317;
   F[3222] := 16.988571;
   F[3223] := 16.988571;
   F[3224] := 17.01389;
   F[3225] := 17.089844;
   F[3226] := 17.158566;
   F[3227] := 17.078993;
   F[3228] := 17.158566;
   F[3229] := 17.122396;
   F[3230] := 17.205584;
   F[3231] := 17.227285;
   F[3232] := 17.24537;
   F[3233] := 17.216434;
   F[3234] := 17.238136;
   F[3235] := 17.31409;
   F[3236] := 17.30324;
   F[3237] := 17.364729;
   F[3238] := 17.346643;
   F[3239] := 17.433449;
   F[3240] := 17.4443;
   F[3241] := 17.415365;
   F[3242] := 17.386429;
   F[3243] := 17.404514;
   F[3244] := 17.45515;
   F[3245] := 17.509403;
   F[3246] := 17.534721;
   F[3247] := 17.574509;
   F[3248] := 17.574509;
   F[3249] := 17.545572;
   F[3250] := 17.603443;
   F[3251] := 17.635996;
   F[3252] := 17.668547;
   F[3253] := 17.730034;
   F[3254] := 17.733652;
   F[3255] := 17.730034;
   F[3256] := 17.766203;
   F[3257] := 17.831308;
   F[3258] := 17.798756;
   F[3259] := 17.849392;
   F[3260] := 17.824074;
   F[3261] := 17.914497;
   F[3262] := 17.892796;
   F[3263] := 17.939816;
   F[3264] := 17.943432;
   F[3265] := 18.00492;
   F[3266] := 18.019386;
   F[3267] := 18.041088;
   F[3268] := 18.055555;
   F[3269] := 18.023003;
   F[3270] := 18.091724;
   F[3271] := 18.149595;
   F[3272] := 18.124277;
   F[3273] := 18.185764;
   F[3274] := 18.214699;
   F[3275] := 18.17853;
   F[3276] := 18.2364;
   F[3277] := 18.258102;
   F[3278] := 18.27257;
   F[3279] := 18.315971;
   F[3280] := 18.315971;
   F[3281] := 18.381077;
   F[3282] := 18.359375;
   F[3283] := 18.370226;
   F[3284] := 18.471498;
   F[3285] := 18.48235;
   F[3286] := 18.467882;
   F[3287] := 18.4932;
   F[3288] := 20.554832;
   F[3289] := 23.021557;
   F[3290] := 25.56062;
   F[3291] := 27.987558;
   F[3292] := 30.50492;
   F[3293] := 33.062065;
   F[3294] := 35.467304;
   F[3295] := 37.94126;
   F[3296] := 40.46224;
   F[3297] := 40.505642;
   F[3298] := 36.4511;
   F[3299] := 32.461662;
   F[3300] := 29.644096;
   F[3301] := 27.083334;
   F[3302] := 24.660011;
   F[3303] := 22.063078;
   F[3304] := 19.632523;
   F[3305] := 17.111546;
   F[3306] := 14.594184;
   F[3307] := 12.149161;
   F[3308] := 9.8307295;
   F[3309] := 9.42202;
   F[3310] := 9.497974;
   F[3311] := 9.436487;
   F[3312] := 9.360533;
   F[3313] := 9.367766;
   F[3314] := 9.302662;
   F[3315] := 9.299046;
   F[3316] := 9.2628765;
   F[3317] := 9.324364;
   F[3318] := 9.230324;
   F[3319] := 9.2628765;
   F[3320] := 9.201389;
   F[3321] := 9.248408;
   F[3322] := 9.161603;
   F[3323] := 9.139901;
   F[3324] := 9.129051;
   F[3325] := 9.129051;
   F[3326] := 9.053096;
   F[3327] := 9.082031;
   F[3328] := 9.038629;
   F[3329] := 9.01331;
   F[3330] := 8.987992;
   F[3331] := 8.95544;
   F[3332] := 8.940972;
   F[3333] := 8.940972;
   F[3334] := 8.9192705;
   F[3335] := 8.904803;
   F[3336] := 8.901186;
   F[3337] := 8.915654;
   F[3338] := 8.828849;
   F[3339] := 8.832465;
   F[3340] := 8.810764;
   F[3341] := 8.79268;
   F[3342] := 8.738426;
   F[3343] := 8.752893;
   F[3344] := 8.749276;
   F[3345] := 8.65162;
   F[3346] := 8.669704;
   F[3347] := 8.65162;
   F[3348] := 8.626302;
   F[3349] := 8.586516;
   F[3350] := 8.633536;
   F[3351] := 8.575665;
   F[3352] := 8.586516;
   F[3353] := 8.5286455;
   F[3354] := 8.470776;
   F[3355] := 8.434607;
   F[3356] := 8.430989;
   F[3357] := 8.478009;
   F[3358] := 8.409288;
   F[3359] := 8.365886;
   F[3360] := 8.33695;
   F[3361] := 8.409288;
   F[3362] := 8.333333;
   F[3363] := 8.344184;
   F[3364] := 8.347801;
   F[3365] := 8.318866;
   F[3366] := 8.322483;
   F[3367] := 8.308015;
   F[3368] := 8.192274;
   F[3369] := 8.250145;
   F[3370] := 8.206742;
   F[3371] := 8.192274;
   F[3372] := 8.163339;
   F[3373] := 8.058449;
   F[3374] := 8.105469;
   F[3375] := 8.112702;
   F[3376] := 8.047599;
   F[3377] := 8.029514;
   F[3378] := 8.080151;
   F[3379] := 8.015046;
   F[3380] := 8.0078125;
   F[3381] := 7.91739;
   F[3382] := 8.015046;
   F[3383] := 7.9318576;
   F[3384] := 7.8956885;
   F[3385] := 7.8993053;
   F[3386] := 7.8667536;
   F[3387] := 7.928241;
   F[3388] := 7.837818;
   F[3389] := 7.9065394;
   F[3390] := 7.7690973;
   F[3391] := 7.837818;
   F[3392] := 7.7907987;
   F[3393] := 7.7437787;
   F[3394] := 7.7437787;
   F[3395] := 7.740162;
   F[3396] := 7.664207;
   F[3397] := 7.7220774;
   F[3398] := 7.635272;
   F[3399] := 7.609954;
   F[3400] := 7.6063366;
   F[3401] := 7.6280384;
   F[3402] := 7.573785;
   F[3403] := 7.5665507;
   F[3404] := 7.5159144;
   F[3405] := 7.5014467;
   F[3406] := 7.4544272;
   F[3407] := 7.5050635;
   F[3408] := 7.4761286;
   F[3409] := 7.425492;
   F[3410] := 7.4399595;
   F[3411] := 7.39294;
   F[3412] := 7.411024;
   F[3413] := 7.385706;
   F[3414] := 7.3350697;
   F[3415] := 7.3350697;
   F[3416] := 7.3386865;
   F[3417] := 7.273582;
   F[3418] := 7.284433;
   F[3419] := 7.2663484;
   F[3420] := 7.2301793;
   F[3421] := 7.2157116;
   F[3422] := 7.1976275;
   F[3423] := 7.157841;
   F[3424] := 7.1940103;
   F[3425] := 7.1867766;
   F[3426] := 7.139757;
   F[3427] := 7.1144385;
   F[3428] := 7.096354;
   F[3429] := 7.081887;
   F[3430] := 7.0638022;
   F[3431] := 7.034867;
   F[3432] := 7.060185;
   F[3433] := 6.9842305;
   F[3434] := 6.854022;
   F[3435] := 6.980613;
   F[3436] := 6.9408274;
   F[3437] := 6.929977;
   F[3438] := 6.904659;
   F[3439] := 6.9118924;
   F[3440] := 6.82147;
   F[3441] := 6.828704;
   F[3442] := 6.817853;
   F[3443] := 6.778067;
   F[3444] := 6.7961516;
   F[3445] := 6.7310476;
   F[3446] := 6.7853007;
   F[3447] := 6.778067;
   F[3448] := 6.702112;
   F[3449] := 6.665943;
   F[3450] := 6.680411;
   F[3451] := 6.629774;
   F[3452] := 6.579138;
   F[3453] := 6.6225405;
   F[3454] := 6.6550927;
   F[3455] := 6.5863714;
   F[3456] := 6.640625;
   F[3457] := 6.5502024;
   F[3458] := 6.5610533;
   F[3459] := 6.514034;
   F[3460] := 6.467014;
   F[3461] := 6.4814816;
   F[3462] := 6.4959493;
   F[3463] := 6.45978;
   F[3464] := 6.430845;
   F[3465] := 6.391059;
   F[3466] := 6.35489;
   F[3467] := 6.391059;
   F[3468] := 6.358507;
   F[3469] := 6.362124;
   F[3470] := 6.35489;
   F[3471] := 6.35489;
   F[3472] := 6.289786;
   F[3473] := 6.25;
   F[3474] := 6.1921296;
   F[3475] := 6.239149;
   F[3476] := 6.221065;
   F[3477] := 6.1921296;
   F[3478] := 6.1704283;
   F[3479] := 6.1306424;
   F[3480] := 6.1631947;
   F[3481] := 6.1306424;
   F[3482] := 6.112558;
   F[3483] := 6.141493;
   F[3484] := 6.069155;
   F[3485] := 6.0149016;
   F[3486] := 6.0257525;
   F[3487] := 6.0149016;
   F[3488] := 5.9136286;
   F[3489] := 5.996817;
   F[3490] := 5.964265;
   F[3491] := 5.920862;
   F[3492] := 5.964265;
   F[3493] := 5.862992;
   F[3494] := 5.9136286;
   F[3495] := 5.870226;
   F[3496] := 5.8521414;
   F[3497] := 5.834057;
   F[3498] := 5.8521414;
   F[3499] := 5.808738;
   F[3500] := 5.794271;
   F[3501] := 5.797888;
   F[3502] := 5.7725697;
   F[3503] := 5.7038484;
   F[3504] := 5.721933;
   F[3505] := 5.6893806;
   F[3506] := 5.6532116;
   F[3507] := 5.721933;
   F[3508] := 5.67853;
   F[3509] := 5.6387444;
   F[3510] := 5.6025753;
   F[3511] := 5.5664062;
   F[3512] := 5.5627894;
   F[3513] := 5.5013022;
   F[3514] := 5.5483217;
   F[3515] := 5.4832177;
   F[3516] := 5.497685;
   F[3517] := 5.497685;
   F[3518] := 5.4615164;
   F[3519] := 5.479601;
   F[3520] := 5.443432;
   F[3521] := 5.4361978;
   F[3522] := 5.392795;
   F[3523] := 5.3819447;
   F[3524] := 5.3710938;
   F[3525] := 5.327691;
   F[3526] := 5.255353;
   F[3527] := 5.3132234;
   F[3528] := 5.2408853;
   F[3529] := 5.186632;
   F[3530] := 5.291522;
   F[3531] := 5.2481194;
   F[3532] := 5.2372684;
   F[3533] := 5.2372684;
   F[3534] := 5.2010994;
   F[3535] := 5.1974826;
   F[3536] := 5.1721644;
   F[3537] := 5.1757812;
   F[3538] := 5.15408;
   F[3539] := 5.15408;
   F[3540] := 5.0962095;
   F[3541] := 4.9153647;
   F[3542] := 4.2426214;
   F[3543] := 3.584346;
   F[3544] := 2.983941;
   F[3545] := 2.3039641;
   F[3546] := 2.0182292;
   F[3547] := 1.9675926;
   F[3548] := 1.9929109;
   F[3549] := 2.0073786;
   F[3550] := 2.0146122;
   F[3551] := 1.9748263;
   F[3552] := 1.9856771;
   F[3553] := 1.9024885;
   F[3554] := 1.9712095;
   F[3555] := 1.8952546;
   F[3556] := 1.9675926;
   F[3557] := 1.9748263;
   F[3558] := 1.9241898;
   F[3559] := 1.9567419;
   F[3560] := 1.9458913;
   F[3561] := 1.9422743;
   F[3562] := 1.9748263;
   F[3563] := 1.8735533;
   F[3564] := 1.9024885;
   F[3565] := 1.9205729;
   F[3566] := 1.9241898;
   F[3567] := 1.9133391;
   F[3568] := 1.880787;
   F[3569] := 1.9350405;
   F[3570] := 1.9567419;
   F[3571] := 1.8590857;
   F[3572] := 1.9024885;
   F[3573] := 1.8880209;
   F[3574] := 1.8373842;
   F[3575] := 1.8590857;
   F[3576] := 1.884404;
   F[3577] := 1.8699363;
   F[3578] := 1.8265336;
   F[3579] := 1.8229166;
   F[3580] := 1.812066;
   F[3581] := 1.8554688;
   F[3582] := 1.8554688;
   F[3583] := 1.848235;
   F[3584] := 1.848235;
   F[3585] := 1.8590857;
   F[3586] := 1.8265336;
   F[3587] := 1.775897;
   F[3588] := 1.8446181;
   F[3589] := 1.8192998;
   F[3590] := 1.7903646;
   F[3591] := 1.8301505;
   F[3592] := 1.8554688;
   F[3593] := 1.7903646;
   F[3594] := 1.739728;
   F[3595] := 1.8012153;
   F[3596] := 1.7614294;
   F[3597] := 1.808449;
   F[3598] := 1.775897;
   F[3599] := 1.7469618;
   F[3600] := 1.7505788;
   F[3601] := 1.8012153;
   F[3602] := 1.7650462;
   F[3603] := 1.7722801;
   F[3604] := 1.7433449;
   F[3605] := 1.775897;
   F[3606] := 2.665654;
   F[3607] := 6.741898;
   F[3608] := 6.904659;
   F[3609] := 6.915509;
   F[3610] := 6.980613;
   F[3611] := 6.9625287;
   F[3612] := 6.8612556;
   F[3613] := 6.958912;
   F[3614] := 6.904659;
   F[3615] := 6.8721066;
   F[3616] := 6.922743;
   F[3617] := 6.9372106;
   F[3618] := 6.929977;
   F[3619] := 6.955295;
   F[3620] := 6.9372106;
   F[3621] := 6.87934;
   F[3622] := 6.904659;
   F[3623] := 6.9625287;
   F[3624] := 6.966146;
   F[3625] := 6.922743;
   F[3626] := 6.9625287;
   F[3627] := 6.92636;
   F[3628] := 6.958912;
   F[3629] := 7.0167823;
   F[3630] := 6.966146;
   F[3631] := 7.071036;
   F[3632] := 6.958912;
   F[3633] := 7.002315;
   F[3634] := 6.969763;
   F[3635] := 6.9769964;
   F[3636] := 6.9842305;
   F[3637] := 7.0131655;
   F[3638] := 7.005932;
   F[3639] := 7.020399;
   F[3640] := 7.0999713;
   F[3641] := 7.067419;
   F[3642] := 7.0384836;
   F[3643] := 7.0240164;
   F[3644] := 7.0167823;
   F[3645] := 7.0384836;
   F[3646] := 7.060185;
   F[3647] := 7.0782695;
   F[3648] := 7.0999713;
   F[3649] := 7.071036;
   F[3650] := 7.139757;
   F[3651] := 7.0891204;
   F[3652] := 7.0384836;
   F[3653] := 7.081887;
   F[3654] := 7.103588;
   F[3655] := 7.1614585;
   F[3656] := 7.1216726;
   F[3657] := 7.1180553;
   F[3658] := 7.092737;
   F[3659] := 7.157841;
   F[3660] := 7.1542244;
   F[3661] := 7.13614;
   F[3662] := 7.1614585;
   F[3663] := 7.107205;
   F[3664] := 7.18316;
   F[3665] := 7.146991;
   F[3666] := 7.2012444;
   F[3667] := 7.1940103;
   F[3668] := 7.1903934;
   F[3669] := 7.107205;
   F[3670] := 7.2012444;
   F[3671] := 7.1506076;
   F[3672] := 7.18316;
   F[3673] := 7.179543;
   F[3674] := 7.1903934;
   F[3675] := 7.1903934;
   F[3676] := 7.233796;
   F[3677] := 7.1940103;
   F[3678] := 7.2012444;
   F[3679] := 7.2157116;
   F[3680] := 7.2012444;
   F[3681] := 7.204861;
   F[3682] := 7.2518806;
   F[3683] := 7.269965;
   F[3684] := 7.2157116;
   F[3685] := 7.2229457;
   F[3686] := 7.244647;
   F[3687] := 7.2916665;
   F[3688] := 7.24103;
   F[3689] := 7.2916665;
   F[3690] := 7.295284;
   F[3691] := 7.295284;
   F[3692] := 7.2627316;
   F[3693] := 7.2518806;
   F[3694] := 7.3025174;
   F[3695] := 7.3025174;
   F[3696] := 7.306134;
   F[3697] := 7.24103;
   F[3698] := 7.2916665;
   F[3699] := 7.313368;
   F[3700] := 7.418258;
   F[3701] := 7.3242188;
   F[3702] := 7.4001737;
   F[3703] := 7.284433;
   F[3704] := 7.349537;
   F[3705] := 7.3386865;
   F[3706] := 7.3278356;
   F[3707] := 7.3784723;
   F[3708] := 7.313368;
   F[3709] := 7.425492;
   F[3710] := 7.3748555;
   F[3711] := 7.3784723;
   F[3712] := 7.4074073;
   F[3713] := 7.3640046;
   F[3714] := 7.418258;
   F[3715] := 7.4291086;
   F[3716] := 7.3640046;
   F[3717] := 7.4001737;
   F[3718] := 7.421875;
   F[3719] := 7.3784723;
   F[3720] := 7.4399595;
   F[3721] := 7.45081;
   F[3722] := 7.4037905;
   F[3723] := 7.4291086;
   F[3724] := 7.4001737;
   F[3725] := 7.4652777;
   F[3726] := 7.4761286;
   F[3727] := 7.458044;
   F[3728] := 7.472512;
   F[3729] := 7.4761286;
   F[3730] := 7.5014467;
   F[3731] := 7.4797454;
   F[3732] := 7.5014467;
   F[3733] := 7.4363427;
   F[3734] := 7.4761286;
   F[3735] := 7.5014467;
   F[3736] := 7.5159144;
   F[3737] := 7.5195312;
   F[3738] := 7.486979;
   F[3739] := 7.526765;
   F[3740] := 7.5448494;
   F[3741] := 7.533999;
   F[3742] := 7.5448494;
   F[3743] := 7.570168;
   F[3744] := 7.5520835;
   F[3745] := 7.548466;
   F[3746] := 7.548466;
   F[3747] := 7.5557003;
   F[3748] := 7.562934;
   F[3749] := 7.559317;
   F[3750] := 7.5810184;
   F[3751] := 7.60272;
   F[3752] := 7.526765;
   F[3753] := 7.5557003;
   F[3754] := 7.595486;
   F[3755] := 7.5882525;
   F[3756] := 7.6533566;
   F[3757] := 7.6171875;
   F[3758] := 7.6171875;
   F[3759] := 7.6425056;
   F[3760] := 7.6497397;
   F[3761] := 7.6280384;
   F[3762] := 7.6497397;
   F[3763] := 7.6533566;
   F[3764] := 7.6822915;
   F[3765] := 7.6533566;
   F[3766] := 7.703993;
   F[3767] := 7.696759;
   F[3768] := 7.70761;
   F[3769] := 7.6822915;
   F[3770] := 7.675058;
   F[3771] := 7.696759;
   F[3772] := 7.7582464;
   F[3773] := 7.7220774;
   F[3774] := 7.6931424;
   F[3775] := 7.7220774;
   F[3776] := 7.7329283;
   F[3777] := 7.7582464;
   F[3778] := 7.7546296;
   F[3779] := 7.7220774;
   F[3780] := 7.7293115;
   F[3781] := 7.7582464;
   F[3782] := 7.7293115;
   F[3783] := 7.761863;
   F[3784] := 7.7437787;
   F[3785] := 7.7256947;
   F[3786] := 7.7582464;
   F[3787] := 7.7980323;
   F[3788] := 7.7944155;
   F[3789] := 7.772714;
   F[3790] := 7.8595195;
   F[3791] := 7.837818;
   F[3792] := 7.8305845;
   F[3793] := 7.7980323;
   F[3794] := 7.877604;
   F[3795] := 7.837818;
   F[3796] := 7.8812213;
   F[3797] := 7.9354744;
   F[3798] := 7.877604;
   F[3799] := 7.921007;
   F[3800] := 7.8812213;
   F[3801] := 7.9029226;
   F[3802] := 7.949942;
   F[3803] := 7.8956885;
   F[3804] := 7.888455;
   F[3805] := 7.921007;
   F[3806] := 7.873987;
   F[3807] := 7.913773;
   F[3808] := 7.8920717;
   F[3809] := 7.924624;
   F[3810] := 7.939091;
   F[3811] := 7.9354744;
   F[3812] := 7.939091;
   F[3813] := 7.9571757;
   F[3814] := 7.949942;
   F[3815] := 7.9716434;
   F[3816] := 7.96441;
   F[3817] := 7.9824944;
   F[3818] := 8.02228;
   F[3819] := 7.993345;
   F[3820] := 8.047599;
   F[3821] := 7.989728;
   F[3822] := 7.986111;
   F[3823] := 8.058449;
   F[3824] := 8.015046;
   F[3825] := 8.087384;
   F[3826] := 7.9788775;
   F[3827] := 8.029514;
   F[3828] := 8.029514;
   F[3829] := 8.015046;
   F[3830] := 8.051215;
   F[3831] := 8.000579;
   F[3832] := 8.065682;
   F[3833] := 8.036748;
   F[3834] := 8.101851;
   F[3835] := 8.130787;
   F[3836] := 8.0910015;
   F[3837] := 8.098235;
   F[3838] := 8.087384;
   F[3839] := 8.109086;
   F[3840] := 8.134404;
   F[3841] := 8.072917;
   F[3842] := 8.130787;
   F[3843] := 8.152489;
   F[3844] := 8.159722;
   F[3845] := 8.159722;
   F[3846] := 8.141638;
   F[3847] := 8.181423;
   F[3848] := 8.152489;
   F[3849] := 8.134404;
   F[3850] := 8.18504;
   F[3851] := 8.156105;
   F[3852] := 8.253761;
   F[3853] := 8.210359;
   F[3854] := 8.206742;
   F[3855] := 8.286314;
   F[3856] := 8.250145;
   F[3857] := 8.264612;
   F[3858] := 8.239294;
   F[3859] := 8.250145;
   F[3860] := 8.264612;
   F[3861] := 8.257379;
   F[3862] := 8.28993;
   F[3863] := 8.28993;
   F[3864] := 8.260995;
   F[3865] := 8.2682295;
   F[3866] := 8.326099;
   F[3867] := 8.3152485;
   F[3868] := 8.39482;
   F[3869] := 8.322483;
   F[3870] := 8.293548;
   F[3871] := 8.297164;
   F[3872] := 8.308015;
   F[3873] := 8.344184;
   F[3874] := 8.369502;
   F[3875] := 8.333333;
   F[3876] := 8.412905;
   F[3877] := 8.39482;
   F[3878] := 8.402055;
   F[3879] := 8.402055;
   F[3880] := 8.467158;
   F[3881] := 8.412905;
   F[3882] := 8.412905;
   F[3883] := 8.420139;
   F[3884] := 8.423756;
   F[3885] := 8.463542;
   F[3886] := 8.456307;
   F[3887] := 8.449074;
   F[3888] := 8.391204;
   F[3889] := 8.53588;
   F[3890] := 8.459925;
   F[3891] := 8.496094;
   F[3892] := 8.48886;
   F[3893] := 8.430989;
   F[3894] := 8.532263;
   F[3895] := 8.510561;
   F[3896] := 8.474392;
   F[3897] := 8.53588;
   F[3898] := 8.525029;
   F[3899] := 8.582899;
   F[3900] := 8.525029;
   F[3901] := 8.532263;
   F[3902] := 8.550347;
   F[3903] := 8.770978;
   F[3904] := 11.060474;
   F[3905] := 13.581452;
   F[3906] := 16.04456;
   F[3907] := 18.518518;
   F[3908] := 21.097366;
   F[3909] := 23.53154;
   F[3910] := 26.016348;
   F[3911] := 28.468605;
   F[3912] := 31.011284;
   F[3913] := 33.52141;
   F[3914] := 35.991753;
   F[3915] := 38.43316;
   F[3916] := 40.91797;
   F[3917] := 40.99754;
   F[3918] := 37.7785;
   F[3919] := 35.380497;
   F[3920] := 32.816116;
   F[3921] := 30.349392;
   F[3922] := 27.81033;
   F[3923] := 25.347221;
   F[3924] := 22.858797;
   F[3925] := 20.413773;
   F[3926] := 17.86386;
   F[3927] := 15.350116;
   F[3928] := 12.91956;
   F[3929] := 10.376881;
   F[3930] := 7.96441;
   F[3931] := 6.8250866;
   F[3932] := 6.8612556;
   F[3933] := 6.8106194;
   F[3934] := 6.8359375;
   F[3935] := 6.8395543;
   F[3936] := 6.8106194;
   F[3937] := 6.792535;
   F[3938] := 6.8106194;
   F[3939] := 6.7744503;
   F[3940] := 6.7853007;
   F[3941] := 6.792535;
   F[3942] := 6.756366;
   F[3943] := 6.7744503;
   F[3944] := 6.7274303;
   F[3945] := 6.7382812;
   F[3946] := 6.756366;
   F[3947] := 6.767216;
   F[3948] := 6.749132;
   F[3949] := 6.6876445;
   F[3950] := 6.7635994;
   F[3951] := 6.7708335;
   F[3952] := 6.7093463;
   F[3953] := 6.702112;
   F[3954] := 6.741898;
   F[3955] := 6.691262;
   F[3956] := 6.640625;
   F[3957] := 6.6948786;
   F[3958] := 6.6333914;
   F[3959] := 6.640625;
   F[3960] := 6.604456;
   F[3961] := 6.651476;
   F[3962] := 6.640625;
   F[3963] := 6.6478586;
   F[3964] := 6.600839;
   F[3965] := 6.5936055;
   F[3966] := 6.6080728;
   F[3967] := 6.5863714;
   F[3968] := 6.5863714;
   F[3969] := 6.6080728;
   F[3970] := 6.6225405;
   F[3971] := 6.6189237;
   F[3972] := 6.579138;
   F[3973] := 6.615307;
   F[3974] := 6.6080728;
   F[3975] := 6.5610533;
   F[3976] := 6.6225405;
   F[3977] := 6.528501;
   F[3978] := 6.5502024;
   F[3979] := 6.524884;
   F[3980] := 6.492332;
   F[3981] := 6.528501;
   F[3982] := 6.5104165;
   F[3983] := 6.532118;
   F[3984] := 6.4453125;
   F[3985] := 6.488715;
   F[3986] := 6.4489293;
   F[3987] := 6.488715;
   F[3988] := 6.4778647;
   F[3989] := 6.4706306;
   F[3990] := 6.463397;
   F[3991] := 6.40191;
   F[3992] := 6.4344616;
   F[3993] := 6.4453125;
   F[3994] := 6.4416957;
   F[3995] := 6.4489293;
   F[3996] := 6.387442;
   F[3997] := 6.4091434;
   F[3998] := 6.423611;
   F[3999] := 6.40191;
   F[4000] := 6.427228;
   F[4001] := 6.427228;
   F[4002] := 6.3946757;
   F[4003] := 6.376591;
   F[4004] := 6.45978;
   F[4005] := 6.3729744;
   F[4006] := 6.351273;
   F[4007] := 6.2970195;
   F[4008] := 6.3838253;
   F[4009] := 6.358507;
   F[4010] := 6.325955;
   F[4011] := 6.3331885;
   F[4012] := 6.289786;
   F[4013] := 6.322338;
   F[4014] := 6.3693576;
   F[4015] := 6.3295717;
   F[4016] := 6.2934027;
   F[4017] := 6.2825522;
   F[4018] := 6.3042536;
   F[4019] := 6.325955;
   F[4020] := 6.184896;
   F[4021] := 6.260851;
   F[4022] := 6.2644677;
   F[4023] := 6.2970195;
   F[4024] := 6.2174478;
   F[4025] := 6.2319155;
   F[4026] := 6.1921296;
   F[4027] := 6.25;
   F[4028] := 6.2427664;
   F[4029] := 6.2029805;
   F[4030] := 6.210214;
   F[4031] := 6.199363;
   F[4032] := 6.239149;
   F[4033] := 6.184896;
   F[4034] := 6.213831;
   F[4035] := 6.1957464;
   F[4036] := 6.1631947;
   F[4037] := 6.239149;
   F[4038] := 6.1559606;
   F[4039] := 6.1559606;
   F[4040] := 6.2065973;
   F[4041] := 6.0872397;
   F[4042] := 6.1668115;
   F[4043] := 6.174045;
   F[4044] := 6.148727;
   F[4045] := 6.101707;
   F[4046] := 6.188513;
   F[4047] := 6.1595774;
   F[4048] := 6.069155;
   F[4049] := 6.148727;
   F[4050] := 6.112558;
   F[4051] := 6.0944734;
   F[4052] := 6.0836225;
   F[4053] := 6.047454;
   F[4054] := 6.0836225;
   F[4055] := 6.061921;
   F[4056] := 6.09809;
   F[4057] := 6.0872397;
   F[4058] := 6.061921;
   F[4059] := 6.1197915;
   F[4060] := 6.0655384;
   F[4061] := 6.061921;
   F[4062] := 6.0185184;
   F[4063] := 6.0944734;
   F[4064] := 6.047454;
   F[4065] := 6.032986;
   F[4066] := 6.04022;
   F[4067] := 6.007668;
   F[4068] := 5.985966;
   F[4069] := 6.007668;
   F[4070] := 6.0221353;
   F[4071] := 5.985966;
   F[4072] := 5.960648;
   F[4073] := 5.996817;
   F[4074] := 5.964265;
   F[4075] := 5.975116;
   F[4076] := 6.0293694;
   F[4077] := 6.0221353;
   F[4078] := 5.9497976;
   F[4079] := 5.9570312;
   F[4080] := 5.964265;
   F[4081] := 6.0040507;
   F[4082] := 5.931713;
   F[4083] := 5.9136286;
   F[4084] := 5.9497976;
   F[4085] := 5.924479;
   F[4086] := 5.9425635;
   F[4087] := 5.9280963;
   F[4088] := 5.9136286;
   F[4089] := 5.8810763;
   F[4090] := 5.870226;
   F[4091] := 5.8810763;
   F[4092] := 5.8412905;
   F[4093] := 5.9280963;
   F[4094] := 5.8449073;
   F[4095] := 5.8449073;
   F[4096] := 5.8774595;
   F[4097] := 5.8376737;
   F[4098] := 5.823206;
   F[4099] := 5.8810763;
   F[4100] := 5.855758;
   F[4101] := 5.855758;
   F[4102] := 5.797888;
   F[4103] := 5.8123555;
   F[4104] := 5.8738427;
   F[4105] := 5.7761865;
   F[4106] := 5.7725697;
   F[4107] := 5.8376737;
   F[4108] := 5.78342;
   F[4109] := 5.743634;
   F[4110] := 5.808738;
   F[4111] := 5.732784;
   F[4112] := 5.8051214;
   F[4113] := 5.7761865;
   F[4114] := 5.747251;
   F[4115] := 5.78342;
   F[4116] := 5.743634;
   F[4117] := 5.8015046;
   F[4118] := 5.743634;
   F[4119] := 5.7364006;
   F[4120] := 5.747251;
   F[4121] := 5.7400174;
   F[4122] := 5.7906537;
   F[4123] := 5.732784;
   F[4124] := 5.671296;
   F[4125] := 5.7400174;
   F[4126] := 5.6640625;
   F[4127] := 5.6893806;
   F[4128] := 5.7038484;
   F[4129] := 5.656829;
   F[4130] := 5.7146993;
   F[4131] := 5.656829;
   F[4132] := 5.649595;
   F[4133] := 5.6640625;
   F[4134] := 5.642361;
   F[4135] := 5.649595;
   F[4136] := 5.711082;
   F[4137] := 5.6676793;
   F[4138] := 5.6893806;
   F[4139] := 5.6604457;
   F[4140] := 5.6315103;
   F[4141] := 5.642361;
   F[4142] := 5.6351275;
   F[4143] := 5.6532116;
   F[4144] := 5.5989585;
   F[4145] := 5.6387444;
   F[4146] := 5.5917244;
   F[4147] := 5.5989585;
   F[4148] := 5.5881076;
   F[4149] := 5.584491;
   F[4150] := 5.617043;
   F[4151] := 5.642361;
   F[4152] := 5.5664062;
   F[4153] := 5.570023;
   F[4154] := 5.5230036;
   F[4155] := 5.62066;
   F[4156] := 5.580874;
   F[4157] := 5.5555553;
   F[4158] := 5.584491;
   F[4159] := 5.5664062;
   F[4160] := 5.544705;
   F[4161] := 5.5374713;
   F[4162] := 5.5555553;
   F[4163] := 5.5266204;
   F[4164] := 5.5374713;
   F[4165] := 5.580874;
   F[4166] := 5.5157695;
   F[4167] := 5.5483217;
   F[4168] := 5.580874;
   F[4169] := 5.497685;
   F[4170] := 5.5013022;
   F[4171] := 5.497685;
   F[4172] := 5.5230036;
   F[4173] := 5.504919;
   F[4174] := 5.497685;
   F[4175] := 5.494068;
   F[4176] := 5.443432;
   F[4177] := 5.504919;
   F[4178] := 5.472367;
   F[4179] := 5.4615164;
   F[4180] := 5.472367;
   F[4181] := 5.4506655;
   F[4182] := 5.457899;
   F[4183] := 5.3855615;
   F[4184] := 5.3493924;
   F[4185] := 5.4144964;
   F[4186] := 5.4217305;
   F[4187] := 5.4217305;
   F[4188] := 5.403646;
   F[4189] := 5.396412;
   F[4190] := 5.3855615;
   F[4191] := 5.428964;
   F[4192] := 5.3855615;
   F[4193] := 5.4253473;
   F[4194] := 5.3819447;
   F[4195] := 5.3819447;
   F[4196] := 5.3240743;
   F[4197] := 5.36386;
   F[4198] := 5.3493924;
   F[4199] := 5.360243;
   F[4200] := 5.3855615;
   F[4201] := 5.353009;
   F[4202] := 5.3891783;
   F[4203] := 5.367477;
   F[4204] := 5.3747106;
   F[4205] := 5.3783274;
   F[4206] := 5.342159;
   F[4207] := 5.3023725;
   F[4208] := 5.3385415;
   F[4209] := 5.2625866;
   F[4210] := 5.266204;
   F[4211] := 5.31684;
   F[4212] := 5.320457;
   F[4213] := 5.3132234;
   F[4214] := 5.367477;
   F[4215] := 5.31684;
   F[4216] := 5.2372684;
   F[4217] := 5.295139;
   F[4218] := 5.2842884;
   F[4219] := 5.2734375;
   F[4220] := 5.251736;
   F[4221] := 5.2698207;
   F[4222] := 5.2698207;
   F[4223] := 5.2010994;
   F[4224] := 5.215567;
   F[4225] := 5.251736;
   F[4226] := 5.215567;
   F[4227] := -0.01808449;
   F[4228] := 2.0688658;
   F[4229] := 2.7307582;
   F[4230] := 3.3600984;
   F[4231] := 3.8519964;
   F[4232] := 3.9134839;
   F[4233] := 3.9026332;
   F[4234] := 3.8953993;
   F[4235] := 3.9171007;
   F[4236] := 3.9568865;
   F[4237] := 3.9568865;
   F[4238] := 3.9858217;
   F[4239] := 4.0039062;
   F[4240] := 4.018374;
   F[4241] := 3.9677372;
   F[4242] := 4.01114;
   F[4243] := 4.007523;
   F[4244] := 4.0509257;
   F[4245] := 4.021991;
   F[4246] := 4.079861;
   F[4247] := 4.184751;
   F[4248] := 4.181134;
   F[4249] := 4.094329;
   F[4250] := 4.1304975;
   F[4251] := 4.1413484;
   F[4252] := 4.191985;
   F[4253] := 4.1739006;
   F[4254] := 4.1775174;
   F[4255] := 4.170284;
   F[4256] := 4.2173033;
   F[4257] := 4.2064524;
   F[4258] := 4.271557;
   F[4259] := 4.2100697;
   F[4260] := 4.195602;
   F[4261] := 4.2896414;
   F[4262] := 4.271557;
   F[4263] := 4.32581;
   F[4264] := 4.307726;
   F[4265] := 4.300492;
   F[4266] := 4.296875;
   F[4267] := 4.333044;
   F[4268] := 4.401765;
   F[4269] := 4.3655963;
   F[4270] := 4.3511286;
   F[4271] := 4.3800635;
   F[4272] := 4.3945312;
   F[4273] := 4.445168;
   F[4274] := 4.434317;
   F[4275] := 4.37283;
   F[4276] := 4.5030384;
   F[4277] := 4.448785;
   F[4278] := 4.4524016;
   F[4279] := 4.5536747;
   F[4280] := 4.510272;
   F[4281] := 4.5645256;
   F[4282] := 4.546441;
   F[4283] := 4.575376;
   F[4284] := 4.575376;
   F[4285] := 4.5970774;
   F[4286] := 4.5645256;
   F[4287] := 4.5898438;
   F[4288] := 4.6296296;
   F[4289] := 4.622396;
   F[4290] := 4.658565;
   F[4291] := 4.6694155;
   F[4292] := 4.626013;
   F[4293] := 4.647714;
   F[4294] := 4.6694155;
   F[4295] := 4.7092013;
   F[4296] := 4.691117;
   F[4297] := 4.7417536;
   F[4298] := 4.7200522;
   F[4299] := 4.7345195;
   F[4300] := 4.814091;
   F[4301] := 4.8104744;
   F[4302] := 4.8828125;
   F[4303] := 4.799624;
   F[4304] := 4.8538775;
   F[4305] := 4.8719616;
   F[4306] := 4.824942;
   F[4307] := 4.9081306;
   F[4308] := 4.8936634;
   F[4309] := 4.951534;
   F[4310] := 4.9442997;
   F[4311] := 4.969618;
   F[4312] := 4.9840856;
   F[4313] := 4.9479165;
   F[4314] := 5.041956;
   F[4315] := 4.9985533;
   F[4316] := 5.027488;
   F[4317] := 5.00217;
   F[4318] := 5.1215277;
   F[4319] := 5.25897;
   F[4320] := 5.356626;
   F[4321] := 5.418113;
   F[4322] := 5.494068;
   F[4323] := 5.5989585;
   F[4324] := 5.6966147;
   F[4325] := 5.78342;
   F[4326] := 5.870226;
   F[4327] := 5.9895835;
   F[4328] := 6.047454;
   F[4329] := 6.188513;
   F[4330] := 6.275318;
   F[4331] := 6.3440394;
   F[4332] := 6.4850984;
   F[4333] := 6.600839;
   F[4334] := 6.6550927;
   F[4335] := 6.749132;
   F[4336] := 6.781684;
   F[4337] := 6.8757234;
   F[4338] := 7.0638022;
   F[4339] := 7.132523;
   F[4340] := 7.2265625;
   F[4341] := 7.2880497;
   F[4342] := 7.360388;
   F[4343] := 7.4797454;
   F[4344] := 7.559317;
   F[4345] := 7.66059;
   F[4346] := 7.7690973;
   F[4347] := 7.863137;
   F[4348] := 7.9716434;
   F[4349] := 8.083767;
   F[4350] := 8.1380205;
   F[4351] := 8.210359;
   F[4352] := 8.358651;
   F[4353] := 8.373119;
   F[4354] := 8.564815;
   F[4355] := 8.666088;
   F[4356] := 8.749276;
   F[4357] := 8.79268;
   F[4358] := 8.940972;
   F[4359] := 9.024161;
   F[4360] := 9.125434;
   F[4361] := 9.205006;
   F[4362] := 9.280961;
   F[4363] := 9.414786;
   F[4364] := 9.501592;
   F[4365] := 9.58478;
   F[4366] := 9.682436;
   F[4367] := 9.740307;
   F[4368] := 8.868634;
   F[4369] := 8.083767;
   F[4370] := 7.269965;
   F[4371] := 6.463397;
   F[4372] := 5.7689524;
   F[4373] := 5.8123555;
   F[4374] := 5.859375;
   F[4375] := 5.855758;
   F[4376] := 5.870226;
   F[4377] := 5.8919272;
   F[4378] := 5.8919272;
   F[4379] := 5.895544;
   F[4380] := 5.975116;
   F[4381] := 6.011285;
   F[4382] := 5.9570312;
   F[4383] := 6.0149016;
   F[4384] := 6.0040507;
   F[4385] := 6.072772;
   F[4386] := 6.076389;
   F[4387] := 6.069155;
   F[4388] := 6.0944734;
   F[4389] := 6.1306424;
   F[4390] := 6.199363;
   F[4391] := 6.1704283;
   F[4392] := 6.1631947;
   F[4393] := 6.184896;
   F[4394] := 6.199363;
   F[4395] := 6.213831;
   F[4396] := 6.2644677;
   F[4397] := 6.2717013;
   F[4398] := 6.3042536;
   F[4399] := 6.322338;
   F[4400] := 6.365741;
   F[4401] := 6.3440394;
   F[4402] := 6.3838253;
   F[4403] := 6.3802085;
   F[4404] := 6.4561634;
   F[4405] := 6.4091434;
   F[4406] := 6.4489293;
   F[4407] := 6.45978;
   F[4408] := 6.528501;
   F[4409] := 6.5067997;
   F[4410] := 6.532118;
   F[4411] := 6.528501;
   F[4412] := 6.589988;
   F[4413] := 6.5936055;
   F[4414] := 6.5719037;
   F[4415] := 6.5936055;
   F[4416] := 6.651476;
   F[4417] := 6.6731772;
   F[4418] := 6.702112;
   F[4419] := 6.712963;
   F[4420] := 6.7201967;
   F[4421] := 6.7093463;
   F[4422] := 6.828704;
   F[4423] := 6.7961516;
   F[4424] := 6.7853007;
   F[4425] := 6.8395543;
   F[4426] := 6.857639;
   F[4427] := 6.8974247;
   F[4428] := 6.8757234;
   F[4429] := 6.919126;
   F[4430] := 6.9516783;
   F[4431] := 6.9335938;
   F[4432] := 6.929977;
   F[4433] := 7.0167823;
   F[4434] := 7.0240164;
   F[4435] := 6.9733796;
   F[4436] := 7.056568;
   F[4437] := 7.042101;
   F[4438] := 7.168692;
   F[4439] := 7.146991;
   F[4440] := 7.1144385;
   F[4441] := 7.143374;
   F[4442] := 7.1650753;
   F[4443] := 7.1506076;
   F[4444] := 7.212095;
   F[4445] := 7.2157116;
   F[4446] := 7.2591147;
   F[4447] := 7.244647;
   F[4448] := 7.2916665;
   F[4449] := 7.309751;
   F[4450] := 7.2916665;
   F[4451] := 7.360388;
   F[4452] := 7.4001737;
   F[4453] := 7.3386865;
   F[4454] := 7.39294;
   F[4455] := 7.4146414;
   F[4456] := 7.4652777;
   F[4457] := 7.4544272;
   F[4458] := 7.483362;
   F[4459] := 7.494213;
   F[4460] := 7.4652777;
   F[4461] := 7.573785;
   F[4462] := 7.631655;
   F[4463] := 7.609954;
   F[4464] := 9.523293;
   F[4465] := 11.97555;
   F[4466] := 14.507379;
   F[4467] := 16.948784;
   F[4468] := 19.509548;
   F[4469] := 21.96904;
   F[4470] := 24.4864;
   F[4471] := 26.938658;
   F[4472] := 29.47772;
   F[4473] := 31.911892;
   F[4474] := 34.3967;
   F[4475] := 36.9647;
   F[4476] := 39.373554;
   F[4477] := 41.858364;
   F[4478] := 41.95602;
   F[4479] := 38.740597;
   F[4480] := 36.295574;
   F[4481] := 33.78183;
   F[4482] := 31.282553;
   F[4483] := 28.725405;
   F[4484] := 26.280382;
   F[4485] := 23.828125;
   F[4486] := 21.296297;
   F[4487] := 18.804253;
   F[4488] := 16.34838;
   F[4489] := 13.841869;
   F[4490] := 11.400463;
   F[4491] := 8.85055;
   F[4492] := 6.4489293;
   F[4493] := 5.9172454;
   F[4494] := 5.870226;
   F[4495] := 5.8521414;
   F[4496] := 5.794271;
   F[4497] := 5.7725697;
   F[4498] := 5.7761865;
   F[4499] := 5.7400174;
   F[4500] := 5.7291665;
   F[4501] := 5.707465;
   F[4502] := 5.6966147;
   F[4503] := 5.671296;
   F[4504] := 5.6676793;
   F[4505] := 5.642361;
   F[4506] := 5.617043;
   F[4507] := 5.6025753;
   F[4508] := 5.577257;
   F[4509] := 5.4868345;
   F[4510] := 5.5555553;
   F[4511] := 5.504919;
   F[4512] := 5.472367;
   F[4513] := 5.4506655;
   F[4514] := 5.439815;
   F[4515] := 5.3891783;
   F[4516] := 5.443432;
   F[4517] := 5.3493924;
   F[4518] := 5.342159;
   F[4519] := 5.360243;
   F[4520] := 5.3819447;
   F[4521] := 5.31684;
   F[4522] := 5.331308;
   F[4523] := 5.295139;
   F[4524] := 5.2842884;
   F[4525] := 5.2336516;
   F[4526] := 5.2336516;
   F[4527] := 5.1757812;
   F[4528] := 5.190249;
   F[4529] := 5.2119503;
   F[4530] := 5.1106772;
   F[4531] := 5.0962095;
   F[4532] := 5.067274;
   F[4533] := 5.10706;
   F[4534] := 5.0564237;
   F[4535] := 5.0600405;
   F[4536] := 4.9877024;
   F[4537] := 5.0094037;
   F[4538] := 4.962384;
   F[4539] := 4.966001;
   F[4540] := 4.962384;
   F[4541] := 4.9189816;
   F[4542] := 4.929832;
   F[4543] := 4.875579;
   F[4544] := 4.904514;
   F[4545] := 4.8430266;
   F[4546] := 4.8466434;
   F[4547] := 4.79239;
   F[4548] := 4.7743053;
   F[4549] := 4.7779226;
   F[4550] := 4.763455;
   F[4551] := 4.712818;
   F[4552] := 4.712818;
   F[4553] := 4.698351;
   F[4554] := 4.6730323;
   F[4555] := 4.6296296;
   F[4556] := 4.6694155;
   F[4557] := 4.636863;
   F[4558] := 4.5934606;
   F[4559] := 4.5572915;
   F[4560] := 4.5898438;
   F[4561] := 4.550058;
   F[4562] := 4.510272;
   F[4563] := 4.513889;
   F[4564] := 4.448785;
   F[4565] := 4.434317;
   F[4566] := 4.448785;
   F[4567] := 4.4162326;
   F[4568] := 4.3836803;
   F[4569] := 4.3438945;
   F[4570] := 4.412616;
   F[4571] := 4.3655963;
   F[4572] := 4.32581;
   F[4573] := 4.322193;
   F[4574] := 4.296875;
   F[4575] := 4.307726;
   F[4576] := 4.2643228;
   F[4577] := 4.2498555;
   F[4578] := 4.260706;
   F[4579] := 4.2136865;
   F[4580] := 4.184751;
   F[4581] := 4.148582;
   F[4582] := 4.1666665;
   F[4583] := 4.1739006;
   F[4584] := 4.0979457;
   F[4585] := 4.0509257;
   F[4586] := 4.1304975;
   F[4587] := 4.11603;
   F[4588] := 4.0400753;
   F[4589] := 4.05816;
   F[4590] := 4.043692;
   F[4591] := 3.9930556;
   F[4592] := 4.0002894;
   F[4593] := 3.9641204;
   F[4594] := 3.9134839;
   F[4595] := 3.9460359;
   F[4596] := 3.9315684;
   F[4597] := 3.8664641;
   F[4598] := 3.8809316;
   F[4599] := 3.8809316;
   F[4600] := 3.8628473;
   F[4601] := 3.870081;
   F[4602] := 3.765191;
   F[4603] := 3.8194444;
   F[4604] := 3.7760417;
   F[4605] := 3.761574;
   F[4606] := 3.7760417;
   F[4607] := 3.7145543;
   F[4608] := 3.7941263;
   F[4609] := 3.7217882;
   F[4610] := 3.768808;
   F[4611] := 3.7181714;
   F[4612] := 3.7109375;
   F[4613] := 3.685619;
   F[4614] := 3.653067;
   F[4615] := 3.6711516;
   F[4616] := 3.6747684;
   F[4617] := 3.6277487;
   F[4618] := 3.5951967;
   F[4619] := 3.653067;
   F[4620] := 3.5807292;
   F[4621] := 3.5771122;
   F[4622] := 3.5662615;
   F[4623] := 3.5879629;
   F[4624] := 3.5373263;
   F[4625] := 3.5264757;
   F[4626] := 3.4939237;
   F[4627] := 3.479456;
   F[4628] := 3.5083911;
   F[4629] := 3.4975405;
   F[4630] := 3.4541378;
   F[4631] := 3.4613714;
   F[4632] := 3.4288194;
   F[4633] := 3.446904;
   F[4634] := 3.3564816;
   F[4635] := 3.4288194;
   F[4636] := 3.414352;
   F[4637] := 3.3854167;
   F[4638] := 3.3926504;
   F[4639] := 3.3311632;
   F[4640] := 3.2769098;
   F[4641] := 3.3962674;
   F[4642] := 3.3275464;
   F[4643] := 3.305845;
   F[4644] := 3.3094618;
   F[4645] := 3.2443576;
   F[4646] := 3.2443576;
   F[4647] := 3.2913773;
   F[4648] := 3.200955;
   F[4649] := 3.1973379;
   F[4650] := 3.2118056;
   F[4651] := 3.193721;
   F[4652] := 3.200955;
   F[4653] := 3.1394675;
   F[4654] := 3.0960648;
   F[4655] := 3.1322339;
   F[4656] := 3.1286168;
   F[4657] := 3.0852141;
   F[4658] := 3.056279;
   F[4659] := 3.0635128;
   F[4660] := 3.0743635;
   F[4661] := 3.0635128;
   F[4662] := 3.0454283;
   F[4663] := 3.0092592;
   F[4664] := 3.0056424;
   F[4665] := 3.0092592;
   F[4666] := 2.9622395;
   F[4667] := 2.9658566;
   F[4668] := 2.980324;
   F[4669] := 2.9730902;
   F[4670] := 2.9333043;
   F[4671] := 2.9333043;
   F[4672] := 2.879051;
   F[4673] := 2.879051;
   F[4674] := 2.879051;
   F[4675] := 2.904369;
   F[4676] := 2.8284144;
   F[4677] := 2.81033;
   F[4678] := 2.7813947;
   F[4679] := 2.8211806;
   F[4680] := 2.8139467;
   F[4681] := 2.879051;
   F[4682] := 2.7596934;
   F[4683] := 2.7633102;
   F[4684] := 2.7271411;
   F[4685] := 2.7596934;
   F[4686] := 2.7090566;
   F[4687] := 2.6909723;
   F[4688] := 2.7235243;
   F[4689] := 2.6439526;
   F[4690] := 2.7162905;
   F[4691] := 2.633102;
   F[4692] := 2.6367188;
   F[4693] := 2.6439526;
   F[4694] := 2.6222513;
   F[4695] := 2.593316;
   F[4696] := 2.5499132;
   F[4697] := 2.6114004;
   F[4698] := 2.5860822;
   F[4699] := 2.5173612;
   F[4700] := 2.5752316;
   F[4701] := 2.4956598;
   F[4702] := 2.4920428;
   F[4703] := 2.5499132;
   F[4704] := 2.4920428;
   F[4705] := 2.4703414;
   F[4706] := 2.481192;
   F[4707] := 2.419705;
   F[4708] := 2.4414062;
   F[4709] := 2.44864;
   F[4710] := 2.3726852;
   F[4711] := 2.4016204;
   F[4712] := 2.419705;
   F[4713] := 2.34375;
   F[4714] := 2.4016204;
   F[4715] := 2.3654513;
   F[4716] := 2.34375;
   F[4717] := 2.3220487;
   F[4718] := 2.307581;
   F[4719] := 2.3148148;
   F[4720] := 2.3003473;
   F[4721] := 2.2967303;
   F[4722] := 2.2822628;
   F[4723] := 2.2243924;
   F[4724] := 2.199074;
   F[4725] := 1.9965278;
   F[4726] := 1.3599538;
   F[4727] := 0.77039933;
   F[4728] := 4.235388;
   F[4729] := 6.915509;
   F[4730] := 6.8323207;
   F[4731] := 6.8865743;
   F[4732] := 6.9082756;
   F[4733] := 6.922743;
   F[4734] := 6.919126;
   F[4735] := 6.9335938;
   F[4736] := 6.922743;
   F[4737] := 6.929977;
   F[4738] := 6.9082756;
   F[4739] := 6.9118924;
   F[4740] := 6.9372106;
   F[4741] := 6.966146;
   F[4742] := 6.9372106;
   F[4743] := 6.966146;
   F[4744] := 6.969763;
   F[4745] := 7.002315;
   F[4746] := 6.969763;
   F[4747] := 6.9733796;
   F[4748] := 6.922743;
   F[4749] := 6.9480615;
   F[4750] := 6.9516783;
   F[4751] := 6.9986978;
   F[4752] := 6.9625287;
   F[4753] := 6.966146;
   F[4754] := 7.0384836;
   F[4755] := 7.0167823;
   F[4756] := 7.0167823;
   F[4757] := 7.060185;
   F[4758] := 6.9769964;
   F[4759] := 7.027633;
   F[4760] := 7.020399;
   F[4761] := 7.042101;
   F[4762] := 7.034867;
   F[4763] := 7.107205;
   F[4764] := 7.0638022;
   F[4765] := 7.0529513;
   F[4766] := 6.995081;
   F[4767] := 7.0638022;
   F[4768] := 7.060185;
   F[4769] := 7.03125;
   F[4770] := 7.0891204;
   F[4771] := 7.1289062;
   F[4772] := 7.0891204;
   F[4773] := 7.0638022;
   F[4774] := 7.0638022;
   F[4775] := 7.042101;
   F[4776] := 7.056568;
   F[4777] := 7.1289062;
   F[4778] := 7.060185;
   F[4779] := 7.132523;
   F[4780] := 7.1144385;
   F[4781] := 7.1216726;
   F[4782] := 7.1216726;
   F[4783] := 7.1650753;
   F[4784] := 7.103588;
   F[4785] := 7.132523;
   F[4786] := 7.1252894;
   F[4787] := 7.1614585;
   F[4788] := 7.13614;
   F[4789] := 7.3423033;
   F[4790] := 7.9824944;
   F[4791] := 8.629919;
   F[4792] := 9.302662;
   F[4793] := 9.993489;
   F[4794] := 10.250289;
   F[4795] := 10.275608;
   F[4796] := 10.239439;
   F[4797] := 10.315393;
   F[4798] := 10.304543;
   F[4799] := 10.362413;
   F[4800] := 10.340712;
   F[4801] := 10.380498;
   F[4802] := 10.441985;
   F[4803] := 10.427517;
   F[4804] := 10.405816;
   F[4805] := 10.449219;
   F[4806] := 10.478154;
   F[4807] := 10.445601;
   F[4808] := 10.499855;
   F[4809] := 10.543258;
   F[4810] := 10.550492;
   F[4811] := 10.550492;
   F[4812] := 10.546875;
   F[4813] := 10.590278;
   F[4814] := 10.619213;
   F[4815] := 10.640914;
   F[4816] := 10.622829;
   F[4817] := 10.619213;
   F[4818] := 10.684318;
   F[4819] := 10.706018;
   F[4820] := 10.745805;
   F[4821] := 10.7421875;
   F[4822] := 10.821759;
   F[4823] := 10.771123;
   F[4824] := 10.767506;
   F[4825] := 10.774739;
   F[4826] := 10.821759;
   F[4827] := 10.8723955;
   F[4828] := 10.883246;
   F[4829] := 10.828993;
   F[4830] := 10.868779;
   F[4831] := 10.876013;
   F[4832] := 10.955585;
   F[4833] := 10.9375;
   F[4834] := 10.912182;
   F[4835] := 10.988136;
   F[4836] := 10.980903;
   F[4837] := 11.053241;
   F[4838] := 11.035156;
   F[4839] := 11.035156;
   F[4840] := 11.020689;
   F[4841] := 11.085793;
   F[4842] := 11.067708;
   F[4843] := 11.111111;
   F[4844] := 11.125579;
   F[4845] := 11.093026;
   F[4846] := 11.176215;
   F[4847] := 11.190682;
   F[4848] := 11.201533;
   F[4849] := 11.212384;
   F[4850] := 11.183449;
   F[4851] := 11.281105;
   F[4852] := 11.295573;
   F[4853] := 11.288339;
   F[4854] := 11.29919;
   F[4855] := 11.338976;
   F[4856] := 11.291956;
   F[4857] := 11.400463;
   F[4858] := 11.433015;
   F[4859] := 11.389612;
   F[4860] := 11.436632;
   F[4861] := 11.41493;
   F[4862] := 11.436632;
   F[4863] := 11.458333;
   F[4864] := 11.487268;
   F[4865] := 11.541522;
   F[4866] := 11.548756;
   F[4867] := 11.581307;
   F[4868] := 11.56684;
   F[4869] := 11.595776;
   F[4870] := 11.588542;
   F[4871] := 11.668114;
   F[4872] := 11.642796;
   F[4873] := 11.631945;
   F[4874] := 11.722367;
   F[4875] := 11.729601;
   F[4876] := 11.689815;
   F[4877] := 11.678964;
   F[4878] := 11.780237;
   F[4879] := 11.76577;
   F[4880] := 11.892361;
   F[4881] := 11.979167;
   F[4882] := 12.051505;
   F[4883] := 12.134693;
   F[4884] := 12.319155;
   F[4885] := 12.322772;
   F[4886] := 12.445746;
   F[4887] := 12.55787;
   F[4888] := 12.659143;
   F[4889] := 12.702546;
   F[4890] := 12.86169;
   F[4891] := 12.973814;
   F[4892] := 13.017217;
   F[4893] := 13.17636;
   F[4894] := 13.259548;
   F[4895] := 13.357204;
   F[4896] := 13.429543;
   F[4897] := 13.603154;
   F[4898] := 13.675492;
   F[4899] := 13.718895;
   F[4900] := 13.809318;
   F[4901] := 14.008246;
   F[4902] := 14.058883;
   F[4903] := 14.152923;
   F[4904] := 14.275897;
   F[4905] := 14.36632;
   F[4906] := 14.438658;
   F[4907] := 14.550781;
   F[4908] := 14.63397;
   F[4909] := 14.713542;
   F[4910] := 14.847367;
   F[4911] := 14.970342;
   F[4912] := 15.006511;
   F[4913] := 15.143952;
   F[4914] := 15.209057;
   F[4915] := 15.3464985;
   F[4916] := 15.476707;
   F[4917] := 15.5598955;
   F[4918] := 15.700954;
   F[4919] := 15.650318;
   F[4920] := 15.878182;
   F[4921] := 15.968605;
   F[4922] := 16.059029;
   F[4923] := 16.109665;
   F[4924] := 16.257957;
   F[4925] := 16.304977;
   F[4926] := 16.489439;
   F[4927] := 16.536459;
   F[4928] := 16.713686;
   F[4929] := 16.749855;
   F[4930] := 16.681135;
   F[4931] := 15.849248;
   F[4932] := 15.04268;
   F[4933] := 14.228877;
   F[4934] := 13.440393;
   F[4935] := 12.879774;
   F[4936] := 12.865307;
   F[4937] := 12.995515;
   F[4938] := 12.962963;
   F[4939] := 12.905092;
   F[4940] := 12.926794;
   F[4941] := 13.013599;
   F[4942] := 13.017217;
   F[4943] := 13.096788;
   F[4944] := 13.035301;
   F[4945] := 13.104022;
   F[4946] := 13.100405;
   F[4947] := 13.1691265;
   F[4948] := 13.190827;
   F[4949] := 13.17636;
   F[4950] := 13.179976;
   F[4951] := 13.212529;
   F[4952] := 13.205296;
   F[4953] := 13.230614;
   F[4954] := 13.263165;
   F[4955] := 13.255932;
   F[4956] := 13.284867;
   F[4957] := 13.306568;
   F[4958] := 13.357204;
   F[4959] := 13.353588;
   F[4960] := 13.317419;
   F[4961] := 13.418693;
   F[4962] := 13.422309;
   F[4963] := 13.451244;
   F[4964] := 13.494647;
   F[4965] := 13.49103;
   F[4966] := 13.5597515;
   F[4967] := 13.53805;
   F[4968] := 13.595921;
   F[4969] := 13.621239;
   F[4970] := 13.624855;
   F[4971] := 13.646557;
   F[4972] := 13.624855;
   F[4973] := 13.697193;
   F[4974] := 13.726129;
   F[4975] := 13.718895;
   F[4976] := 13.7369795;
   F[4977] := 13.762298;
   F[4978] := 13.798467;
   F[4979] := 13.751447;
   F[4980] := 13.838252;
   F[4981] := 13.812934;
   F[4982] := 13.86357;
   F[4983] := 13.903357;
   F[4984] := 13.870805;
   F[4985] := 13.986546;
   F[4986] := 13.972077;
   F[4987] := 13.935908;
   F[4988] := 14.019097;
   F[4989] := 14.044415;
   F[4990] := 14.0625;
   F[4991] := 14.1276045;
   F[4992] := 14.076967;
   F[4993] := 14.102286;
   F[4994] := 14.080585;
   F[4995] := 14.145689;
   F[4996] := 14.163774;
   F[4997] := 14.196325;
   F[4998] := 14.243345;
   F[4999] := 14.26143;
   F[5000] := 14.268663;
   F[5001] := 14.293982;
   F[5002] := 14.308449;
   F[5003] := 14.315682;
   F[5004] := 14.359086;
   F[5005] := 14.384404;
   F[5006] := 14.3880205;
   F[5007] := 14.637587;
   F[5008] := 17.12963;
   F[5009] := 19.545717;
   F[5010] := 22.106482;
   F[5011] := 24.594908;
   F[5012] := 27.02908;
   F[5013] := 29.542824;
   F[5014] := 32.00955;
   F[5015] := 34.49074;
   F[5016] := 37.01172;
   F[5017] := 39.50376;
   F[5018] := 41.923466;
   F[5019] := 41.927082;
   F[5020] := 38.925056;
   F[5021] := 36.342594;
   F[5022] := 33.778214;
   F[5023] := 31.369358;
   F[5024] := 28.884548;
   F[5025] := 26.425058;
   F[5026] := 23.969185;
   F[5027] := 21.45544;
   F[5028] := 18.927229;
   F[5029] := 16.536459;
   F[5030] := 14.026331;
   F[5031] := 12.742332;
   F[5032] := 12.666377;
   F[5033] := 12.641059;
   F[5034] := 12.684462;
   F[5035] := 12.572338;
   F[5036] := 12.579572;
   F[5037] := 12.594039;
   F[5038] := 12.514467;
   F[5039] := 12.478298;
   F[5040] := 12.471065;
   F[5041] := 12.521702;
   F[5042] := 12.416811;
   F[5043] := 12.413195;
   F[5044] := 12.3878765;
   F[5045] := 12.416811;
   F[5046] := 12.351707;
   F[5047] := 12.319155;
   F[5048] := 12.333623;
   F[5049] := 12.333623;
   F[5050] := 12.275752;
   F[5051] := 12.286603;
   F[5052] := 12.297454;
   F[5053] := 12.188947;
   F[5054] := 12.185329;
   F[5055] := 12.188947;
   F[5056] := 12.1744795;
   F[5057] := 12.185329;
   F[5058] := 12.160011;
   F[5059] := 12.073206;
   F[5060] := 12.112992;
   F[5061] := 12.069589;
   F[5062] := 12.069589;
   F[5063] := 11.968316;
   F[5064] := 12.037037;
   F[5065] := 11.942998;
   F[5066] := 11.924913;
   F[5067] := 11.903212;
   F[5068] := 11.877893;
   F[5069] := 11.895978;
   F[5070] := 11.885127;
   F[5071] := 11.877893;
   F[5072] := 11.798322;
   F[5073] := 11.780237;
   F[5074] := 11.736835;
   F[5075] := 11.77662;
   F[5076] := 11.736835;
   F[5077] := 11.682581;
   F[5078] := 11.668114;
   F[5079] := 11.689815;
   F[5080] := 11.646412;
   F[5081] := 11.6536455;
   F[5082] := 11.621094;
   F[5083] := 11.574074;
   F[5084] := 11.61386;
   F[5085] := 11.490886;
   F[5086] := 11.541522;
   F[5087] := 11.548756;
   F[5088] := 11.443866;
   F[5089] := 11.505353;
   F[5090] := 11.469184;
   F[5091] := 11.436632;
   F[5092] := 11.3932295;
   F[5093] := 11.371528;
   F[5094] := 11.3932295;
   F[5095] := 11.338976;
   F[5096] := 11.313658;
   F[5097] := 11.291956;
   F[5098] := 11.248553;
   F[5099] := 11.266638;
   F[5100] := 11.244936;
   F[5101] := 11.244936;
   F[5102] := 11.1943;
   F[5103] := 11.190682;
   F[5104] := 11.205151;
   F[5105] := 11.201533;
   F[5106] := 11.129195;
   F[5107] := 11.121962;
   F[5108] := 11.107494;
   F[5109] := 11.093026;
   F[5110] := 11.027923;
   F[5111] := 11.064092;
   F[5112] := 11.046007;
   F[5113] := 11.020689;
   F[5114] := 10.99537;
   F[5115] := 10.966435;
   F[5116] := 10.933883;
   F[5117] := 10.926649;
   F[5118] := 10.87963;
   F[5119] := 10.883246;
   F[5120] := 10.792824;
   F[5121] := 10.839844;
   F[5122] := 10.854311;
   F[5123] := 10.839844;
   F[5124] := 10.767506;
   F[5125] := 10.763889;
   F[5126] := 10.724103;
   F[5127] := 10.760272;
   F[5128] := 10.716869;
   F[5129] := 10.698785;
   F[5130] := 10.651765;
   F[5131] := 10.673467;
   F[5132] := 10.662616;
   F[5133] := 10.630064;
   F[5134] := 10.615596;
   F[5135] := 10.637298;
   F[5136] := 10.539641;
   F[5137] := 10.561342;
   F[5138] := 10.492621;
   F[5139] := 10.514323;
   F[5140] := 10.420283;
   F[5141] := 10.441985;
   F[5142] := 10.449219;
   F[5143] := 10.445601;
   F[5144] := 10.384114;
   F[5145] := 10.394965;
   F[5146] := 10.391349;
   F[5147] := 10.340712;
   F[5148] := 10.300926;
   F[5149] := 10.286458;
   F[5150] := 10.250289;
   F[5151] := 10.340712;
   F[5152] := 10.243055;
   F[5153] := 10.250289;
   F[5154] := 10.196036;
   F[5155] := 10.192419;
   F[5156] := 10.177952;
   F[5157] := 10.152633;
   F[5158] := 10.145399;
   F[5159] := 10.163484;
   F[5160] := 10.105614;
   F[5161] := 10.054976;
   F[5162] := 10.069445;
   F[5163] := 10.047743;
   F[5164] := 9.968171;
   F[5165] := 10.062211;
   F[5166] := 9.979022;
   F[5167] := 10.00434;
   F[5168] := 9.997107;
   F[5169] := 9.964555;
   F[5170] := 9.932002;
   F[5171] := 9.892217;
   F[5172] := 9.924768;
   F[5173] := 9.866899;
   F[5174] := 9.8307295;
   F[5175] := 9.812645;
   F[5176] := 9.765625;
   F[5177] := 9.743923;
   F[5178] := 9.780092;
   F[5179] := 9.751158;
   F[5180] := 9.74754;
   F[5181] := 9.704138;
   F[5182] := 9.628182;
   F[5183] := 9.689671;
   F[5184] := 9.660735;
   F[5185] := 9.613715;
   F[5186] := 9.635417;
   F[5187] := 9.620949;
   F[5188] := 9.559462;
   F[5189] := 9.516059;
   F[5190] := 9.544994;
   F[5191] := 9.606482;
   F[5192] := 9.483507;
   F[5193] := 9.505208;
   F[5194] := 9.447338;
   F[5195] := 9.490741;
   F[5196] := 9.4401045;
   F[5197] := 9.436487;
   F[5198] := 9.382234;
   F[5199] := 9.403935;
   F[5200] := 9.382234;
   F[5201] := 9.371383;
   F[5202] := 9.331597;
   F[5203] := 9.31713;
   F[5204] := 9.27011;
   F[5205] := 9.306279;
   F[5206] := 9.248408;
   F[5207] := 9.259259;
   F[5208] := 9.27011;
   F[5209] := 9.172454;
   F[5210] := 9.143518;
   F[5211] := 9.139901;
   F[5212] := 9.1796875;
   F[5213] := 9.129051;
   F[5214] := 9.089265;
   F[5215] := 9.078414;
   F[5216] := 9.092882;
   F[5217] := 9.078414;
   F[5218] := 9.01331;
   F[5219] := 9.0494795;
   F[5220] := 8.973524;
   F[5221] := 8.980758;
   F[5222] := 9.024161;
   F[5223] := 8.959057;
   F[5224] := 9.00246;
   F[5225] := 8.908421;
   F[5226] := 8.857783;
   F[5227] := 8.861401;
   F[5228] := 8.854167;
   F[5229] := 8.80353;
   F[5230] := 8.861401;
   F[5231] := 8.760127;
   F[5232] := 8.85055;
   F[5233] := 8.817998;
   F[5234] := 8.734809;
   F[5235] := 8.731193;
   F[5236] := 8.702257;
   F[5237] := 8.723958;
   F[5238] := 8.734809;
   F[5239] := 8.6588545;
   F[5240] := 8.619068;
   F[5241] := 8.615452;
   F[5242] := 8.608217;
   F[5243] := 8.579283;
   F[5244] := 8.503327;
   F[5245] := 7.8559027;
   F[5246] := 7.309751;
   F[5247] := 6.6333914;
   F[5248] := 5.964265;
   F[5249] := 5.530237;
   F[5250] := 5.541088;
   F[5251] := 5.5121527;
   F[5252] := 5.4759836;
   F[5253] := 5.533854;
   F[5254] := 5.5013022;
   F[5255] := 5.494068;
   F[5256] := 5.5013022;
   F[5257] := 5.5157695;
   F[5258] := 5.3855615;
   F[5259] := 5.4470487;
   F[5260] := 5.439815;
   F[5261] := 5.544705;
   F[5262] := 5.4615164;
   F[5263] := 5.443432;
   F[5264] := 5.360243;
   F[5265] := 5.4000287;
   F[5266] := 5.432581;
   F[5267] := 5.4000287;
   F[5268] := 5.367477;
   F[5269] := 5.4470487;
   F[5270] := 5.3710938;
   F[5271] := 5.4253473;
   F[5272] := 5.3783274;
   F[5273] := 5.396412;
   F[5274] := 5.4470487;
   F[5275] := 5.3240743;
   F[5276] := 5.3710938;
   F[5277] := 5.4108796;
   F[5278] := 5.4361978;
   F[5279] := 5.342159;
   F[5280] := 5.353009;
   F[5281] := 5.367477;
   F[5282] := 5.4000287;
   F[5283] := 5.392795;
   F[5284] := 5.4108796;
   F[5285] := 5.3059897;
   F[5286] := 5.331308;
   F[5287] := 5.3710938;
   F[5288] := 5.31684;
   F[5289] := 5.360243;
   F[5290] := 5.327691;
   F[5291] := 5.327691;
   F[5292] := 5.31684;
   F[5293] := 5.287905;
   F[5294] := 5.2228007;
   F[5295] := 5.3493924;
   F[5296] := 5.331308;
   F[5297] := 5.2987556;
   F[5298] := 5.255353;
   F[5299] := 5.3096066;
   F[5300] := 5.287905;
   F[5301] := 5.266204;
   F[5302] := 5.266204;
   F[5303] := 5.2119503;
   F[5304] := 5.2228007;
   F[5305] := 5.2408853;
   F[5306] := 5.2842884;
   F[5307] := 5.230035;
   F[5308] := 5.1974826;
   F[5309] := -0.047019675;
   F[5310] := 1.5661169;
   F[5311] := 5.5266204;
   F[5312] := 6.0583043;
   F[5313] := 6.0908566;
   F[5314] := 6.0583043;
   F[5315] := 6.141493;
   F[5316] := 6.1161747;
   F[5317] := 6.069155;
   F[5318] := 6.1631947;
   F[5319] := 6.076389;
   F[5320] := 6.101707;
   F[5321] := 6.141493;
   F[5322] := 6.1559606;
   F[5323] := 6.1595774;
   F[5324] := 6.112558;
   F[5325] := 6.1523438;
   F[5326] := 6.141493;
   F[5327] := 6.076389;
   F[5328] := 6.2065973;
   F[5329] := 6.1270256;
   F[5330] := 6.1053243;
   F[5331] := 6.101707;
   F[5332] := 6.1921296;
   F[5333] := 6.137876;
   F[5334] := 6.1812787;
   F[5335] := 6.137876;
   F[5336] := 6.174045;
   F[5337] := 6.1921296;
   F[5338] := 6.2282987;
   F[5339] := 6.260851;
   F[5340] := 6.174045;
   F[5341] := 6.260851;
   F[5342] := 6.174045;
   F[5343] := 6.2065973;
   F[5344] := 6.224682;
   F[5345] := 6.2427664;
   F[5346] := 6.246383;
   F[5347] := 6.2572336;
   F[5348] := 6.289786;
   F[5349] := 6.224682;
   F[5350] := 6.246383;
   F[5351] := 6.1812787;
   F[5352] := 6.2825522;
   F[5353] := 6.213831;
   F[5354] := 6.239149;
   F[5355] := 6.224682;
   F[5356] := 6.260851;
   F[5357] := 6.2680845;
   F[5358] := 6.2680845;
   F[5359] := 6.3042536;
   F[5360] := 6.253617;
   F[5361] := 6.2572336;
   F[5362] := 6.3295717;
   F[5363] := 6.246383;
   F[5364] := 6.3187213;
   F[5365] := 6.3404226;
   F[5366] := 6.3404226;
   F[5367] := 6.311487;
   F[5368] := 6.2717013;
   F[5369] := 6.325955;
   F[5370] := 6.286169;
   F[5371] := 6.278935;
   F[5372] := 6.87934;
   F[5373] := 7.494213;
   F[5374] := 8.11632;
   F[5375] := 8.828849;
   F[5376] := 9.371383;
   F[5377] := 9.414786;
   F[5378] := 9.461805;
   F[5379] := 9.505208;
   F[5380] := 9.483507;
   F[5381] := 9.461805;
   F[5382] := 9.566695;
   F[5383] := 9.476274;
   F[5384] := 9.566695;
   F[5385] := 9.592014;
   F[5386] := 9.58478;
   F[5387] := 9.642651;
   F[5388] := 9.58478;
   F[5389] := 9.689671;
   F[5390] := 9.711371;
   F[5391] := 9.671586;
   F[5392] := 9.67882;
   F[5393] := 9.646267;
   F[5394] := 9.696904;
   F[5395] := 9.74754;
   F[5396] := 9.790943;
   F[5397] := 9.787327;
   F[5398] := 9.812645;
   F[5399] := 9.85243;
   F[5400] := 9.841579;
   F[5401] := 9.863281;
   F[5402] := 9.866899;
   F[5403] := 9.89945;
   F[5404] := 9.884983;
   F[5405] := 9.950087;
   F[5406] := 9.953704;
   F[5407] := 9.997107;
   F[5408] := 9.979022;
   F[5409] := 9.993489;
   F[5410] := 10.047743;
   F[5411] := 10.0441265;
   F[5412] := 10.105614;
   F[5413] := 10.116464;
   F[5414] := 10.076678;
   F[5415] := 10.047743;
   F[5416] := 10.09838;
   F[5417] := 10.101996;
   F[5418] := 10.145399;
   F[5419] := 10.196036;
   F[5420] := 10.239439;
   F[5421] := 10.199653;
   F[5422] := 10.206886;
   F[5423] := 10.246673;
   F[5424] := 10.311776;
   F[5425] := 10.279224;
   F[5426] := 10.293693;
   F[5427] := 10.311776;
   F[5428] := 10.319011;
   F[5429] := 10.358796;
   F[5430] := 10.398582;
   F[5431] := 10.380498;
   F[5432] := 10.441985;
   F[5433] := 10.402199;
   F[5434] := 10.4817705;
   F[5435] := 10.409432;
   F[5436] := 10.478154;
   F[5437] := 10.445601;
   F[5438] := 10.590278;
   F[5439] := 10.507089;
   F[5440] := 10.590278;
   F[5441] := 10.536024;
   F[5442] := 10.56496;
   F[5443] := 10.583044;
   F[5444] := 10.648149;
   F[5445] := 10.608362;
   F[5446] := 10.695168;
   F[5447] := 10.6807;
   F[5448] := 10.698785;
   F[5449] := 10.771123;
   F[5450] := 10.716869;
   F[5451] := 10.807292;
   F[5452] := 10.756655;
   F[5453] := 10.818142;
   F[5454] := 10.8253765;
   F[5455] := 10.8723955;
   F[5456] := 10.814526;
   F[5457] := 10.915798;
   F[5458] := 10.886864;
   F[5459] := 10.962818;
   F[5460] := 10.933883;
   F[5461] := 10.9375;
   F[5462] := 11.024305;
   F[5463] := 11.08941;
   F[5464] := 11.168982;
   F[5465] := 11.273871;
   F[5466] := 11.422164;
   F[5467] := 11.487268;
   F[5468] := 11.577691;
   F[5469] := 11.66088;
   F[5470] := 11.791088;
   F[5471] := 11.942998;
   F[5472] := 12.004485;
   F[5473] := 12.051505;
   F[5474] := 12.116609;
   F[5475] := 12.2432;
   F[5476] := 12.380642;
   F[5477] := 12.449364;
   F[5478] := 12.597656;
   F[5479] := 12.680845;
   F[5480] := 12.764033;
   F[5481] := 12.847222;
   F[5482] := 12.948495;
   F[5483] := 13.064236;
   F[5484] := 13.147425;
   F[5485] := 13.245081;
   F[5486] := 13.378906;
   F[5487] := 13.418693;
   F[5488] := 13.610388;
   F[5489] := 13.646557;
   F[5490] := 13.70081;
   F[5491] := 13.8671875;
   F[5492] := 13.925057;
   F[5493] := 14.087818;
   F[5494] := 14.160156;
   F[5495] := 14.275897;
   F[5496] := 14.355469;
   F[5497] := 14.43504;
   F[5498] := 14.510995;
   F[5499] := 14.680989;
   F[5500] := 14.756945;
   F[5501] := 14.832899;
   F[5502] := 14.966724;
   F[5503] := 15.046296;
   F[5504] := 15.154803;
   F[5505] := 15.292245;
   F[5506] := 15.389901;
   F[5507] := 15.455006;
   F[5508] := 15.5598955;
   F[5509] := 15.628617;
   F[5510] := 15.794994;
   F[5511] := 15.867332;
   F[5512] := 15.954138;
   F[5513] := 15.353733;
   F[5514] := 14.612268;
   F[5515] := 13.7839985;
   F[5516] := 13.0027485;
   F[5517] := 12.123842;
   F[5518] := 12.076823;
   F[5519] := 12.087673;
   F[5520] := 12.094908;
   F[5521] := 12.09129;
   F[5522] := 12.120226;
   F[5523] := 12.203414;
   F[5524] := 12.178096;
   F[5525] := 12.160011;
   F[5526] := 12.203414;
   F[5527] := 12.250434;
   F[5528] := 12.268518;
   F[5529] := 12.311921;
   F[5530] := 12.3046875;
   F[5531] := 12.3046875;
   F[5532] := 12.340857;
   F[5533] := 12.337239;
   F[5534] := 12.380642;
   F[5535] := 12.398726;
   F[5536] := 12.416811;
   F[5537] := 12.481915;
   F[5538] := 12.492766;
   F[5539] := 12.528935;
   F[5540] := 12.460214;
   F[5541] := 12.525318;
   F[5542] := 12.518085;
   F[5543] := 12.561487;
   F[5544] := 12.550636;
   F[5545] := 12.572338;
   F[5546] := 12.644676;
   F[5547] := 12.662761;
   F[5548] := 12.69893;
   F[5549] := 12.706163;
   F[5550] := 12.720631;
   F[5551] := 12.70978;
   F[5552] := 12.745949;
   F[5553] := 12.771267;
   F[5554] := 12.767651;
   F[5555] := 12.843605;
   F[5556] := 12.8255205;
   F[5557] := 12.86169;
   F[5558] := 12.87254;
   F[5559] := 12.879774;
   F[5560] := 12.944879;
   F[5561] := 12.966579;
   F[5562] := 12.915943;
   F[5563] := 12.962963;
   F[5564] := 12.97743;
   F[5565] := 13.042535;
   F[5566] := 13.053386;
   F[5567] := 13.107639;
   F[5568] := 13.118489;
   F[5569] := 13.132957;
   F[5570] := 13.1691265;
   F[5571] := 13.12934;
   F[5572] := 13.198061;
   F[5573] := 13.194445;
   F[5574] := 13.248698;
   F[5575] := 13.263165;
   F[5576] := 13.274016;
   F[5577] := 13.292101;
   F[5578] := 13.321036;
   F[5579] := 13.342737;
   F[5580] := 13.3463545;
   F[5581] := 13.411458;
   F[5582] := 13.389757;
   F[5583] := 13.425926;
   F[5584] := 13.43316;
   F[5585] := 13.483796;
   F[5586] := 13.530816;
   F[5587] := 13.512732;
   F[5588] := 13.556134;
   F[5589] := 13.545283;
   F[5590] := 13.563368;
   F[5591] := 13.603154;
   F[5592] := 13.6067705;
   F[5593] := 13.697193;
   F[5594] := 13.671875;
   F[5595] := 13.715278;
   F[5596] := 13.722511;
   F[5597] := 13.733362;
   F[5598] := 13.762298;
   F[5599] := 13.827401;
   F[5600] := 13.776765;
   F[5601] := 13.859954;
   F[5602] := 13.870805;
   F[5603] := 13.899739;
   F[5604] := 13.914207;
   F[5605] := 13.91059;
   F[5606] := 13.943142;
   F[5607] := 13.91059;
   F[5608] := 14.001013;
   F[5609] := 14.9088545;
   F[5610] := 17.379196;
   F[5611] := 19.874855;
   F[5612] := 22.363281;
   F[5613] := 24.927662;
   F[5614] := 27.434172;
   F[5615] := 29.868345;
   F[5616] := 32.37124;
   F[5617] := 34.84158;
   F[5618] := 37.351707;
   F[5619] := 39.850983;
   F[5620] := 42.30324;
   F[5621] := 42.317707;
   F[5622] := 38.404224;
   F[5623] := 35.919415;
   F[5624] := 33.412907;
   F[5625] := 30.917246;
   F[5626] := 28.464989;
   F[5627] := 25.951244;
   F[5628] := 23.441116;
   F[5629] := 20.916521;
   F[5630] := 18.478733;
   F[5631] := 15.9505205;
   F[5632] := 13.469329;
   F[5633] := 11.038774;
   F[5634] := 10.152633;
   F[5635] := 10.141783;
   F[5636] := 10.0911455;
   F[5637] := 10.087529;
   F[5638] := 10.101996;
   F[5639] := 10.058594;
   F[5640] := 10.033276;
   F[5641] := 10.00434;
   F[5642] := 9.997107;
   F[5643] := 9.89945;
   F[5644] := 9.950087;
   F[5645] := 9.950087;
   F[5646] := 9.942853;
   F[5647] := 9.870515;
   F[5648] := 9.845197;
   F[5649] := 9.801794;
   F[5650] := 9.8307295;
   F[5651] := 9.798177;
   F[5652] := 9.790943;
   F[5653] := 9.790943;
   F[5654] := 9.725839;
   F[5655] := 9.664351;
   F[5656] := 9.7005205;
   F[5657] := 9.704138;
   F[5658] := 9.624566;
   F[5659] := 9.664351;
   F[5660] := 9.58478;
   F[5661] := 9.559462;
   F[5662] := 9.563079;
   F[5663] := 9.544994;
   F[5664] := 9.512443;
   F[5665] := 9.541377;
   F[5666] := 9.4871235;
   F[5667] := 9.454572;
   F[5668] := 9.425636;
   F[5669] := 9.447338;
   F[5670] := 9.396702;
   F[5671] := 9.382234;
   F[5672] := 9.360533;
   F[5673] := 9.346065;
   F[5674] := 9.342448;
   F[5675] := 9.331597;
   F[5676] := 9.3098955;
   F[5677] := 9.288195;
   F[5678] := 9.212239;
   F[5679] := 9.241175;
   F[5680] := 9.172454;
   F[5681] := 9.215857;
   F[5682] := 9.168837;
   F[5683] := 9.154369;
   F[5684] := 9.132668;
   F[5685] := 9.092882;
   F[5686] := 9.027778;
   F[5687] := 9.092882;
   F[5688] := 9.024161;
   F[5689] := 8.984375;
   F[5690] := 8.987992;
   F[5691] := 8.948206;
   F[5692] := 8.908421;
   F[5693] := 8.937355;
   F[5694] := 8.875868;
   F[5695] := 8.893952;
   F[5696] := 8.861401;
   F[5697] := 8.854167;
   F[5698] := 8.828849;
   F[5699] := 8.832465;
   F[5700] := 8.817998;
   F[5701] := 8.756511;
